FUNCTION_BLOCK FB_CIP EXTENDS FB_SFC_Cycle IMPLEMENTS ITF_FB_SFC_Cycle
VAR_INPUT
	valFillWater_T91	: E_Pis_Name;
	valFillWater_T92	: E_Pis_Name;
	valFillWater_T93	: E_Pis_Name;
	valFillWater_T94	: E_Pis_Name;
	
	lvlTank_T91			: ST_Tank_Level	;
	lvlTank_T92			: ST_Tank_Level	;
	lvlTank_T93			: ST_Tank_Level	;
	lvlTank_T94			: ST_Tank_Level	;

END_VAR
VAR_OUTPUT
END_VAR
VAR
	//bRun: BOOL;
	eRun: E_CIP_Source;

	eMode			: E_CIP_Mode;
	eCIP_Return		: E_CIP_Return;
	eCIP_Source		: E_CIP_Source;
	eCIP_Usage		: E_CIP_Usage;
	eReq			: ST_CIP_Request;
	eReqBlank		: ST_CIP_Request;
	eReqLocal		: ST_CIP_Request;
	
	ref_lvlTank_Client		: REFERENCE TO ST_Tank_Level	;

	//bStepDone: BOOL;
	
	iPosSelect_HMI: INT;

	rtPosMoveHMI_Up		: R_TRIG;
	rtPosMoveHMI_Down	: R_TRIG;
	rtPosDeleteHMI		: R_TRIG;
	rtPosDeleteAllHMI	: R_TRIG;
	
	eRefClient_fbElement		: REFERENCE TO FB_Element; // FB_Element // E_Element_State_Long
	bClientRef_done				: BOOL;
	fbElement_Blank				: FB_Element;
	eState_Long_Blank			: E_Element_State_Long;
	
	fbPis						: FB_Piston;
	stPis_FillWater_T91			: REFERENCE TO ST_Piston;
	stPis_FillWater_T92			: REFERENCE TO ST_Piston;
	stPis_FillWater_T93			: REFERENCE TO ST_Piston;
	stPis_FillWater_T94			: REFERENCE TO ST_Piston;
	
	rtReqLocalCIP_Full_HMI: R_TRIG;
	rtReqLocalCIP_Detergent_HMI: R_TRIG;
	rtReqCleanEmpty_HMI: R_TRIG;
	rtModeOff: R_TRIG;
	rtModeManual: R_TRIG;
	rtModeAuto: R_TRIG;
	bTemp: BOOL;
		
	//Process Control
	//concentration
	stDetergent					:	REFERENCE TO ST_ProcessControl	;
	pcDetergent					: 	REFERENCE TO FB_ProcessControl	;	//detergent local
	stDisInfectant				:	REFERENCE TO ST_ProcessControl	;
	pcDisInfectant				: 	REFERENCE TO FB_ProcessControl	;	//detergent local
    //temperature
	stHeatExchanger					:	REFERENCE TO ST_ProcessControl	;
	pcHeatExchanger					: 	REFERENCE TO FB_ProcessControl	;	//	
	stTemperature_Deterg			:	REFERENCE TO ST_ProcessControl	;
	pcTemperature_Deterg			: 	REFERENCE TO FB_ProcessControl	;	//detergent Client	
	stTemperature_Dis				:	REFERENCE TO ST_ProcessControl	;
	pcTemperature_Dis				: 	REFERENCE TO FB_ProcessControl	;//disinfectant local/client
	//temperature client return
	stTemp_ClntReturn				:	REFERENCE TO ST_ProcessControl	;//Client return temperature
	pcTemp_ClntReturn				: 	REFERENCE TO FB_ProcessControl	;//Client return temperature
	
	//flow rate
	stFlow1_Rate					:	REFERENCE TO ST_ProcessControl	;//CIP
	pcFlow1_Rate					: 	REFERENCE TO FB_ProcessControl	;//disinfectant local/client
	stFlow2_Rate					:	REFERENCE TO ST_ProcessControl	;//CIP send
	pcFlow2_Rate					: 	REFERENCE TO FB_ProcessControl	;//disinfectant local/client	return 
	stFlow3_Rate					:	REFERENCE TO ST_ProcessControl	;//CIP send
	pcFlow3_Rate					: 	REFERENCE TO FB_ProcessControl	;//disinfectant local/client	return 
	
	stColor_Level					:	REFERENCE TO ST_ProcessControl	;//CLient CIP //level control 
	pcColor_Level					: 	REFERENCE TO FB_ProcessControl	;//disinfectant local/client //level control 
	stMarinada_Level				:	REFERENCE TO ST_ProcessControl	;//CLient CIP //level control 
	pcMarinada_Level				: 	REFERENCE TO FB_ProcessControl	;//disinfectant local/client //level control 
	
	
	//colar marinade 
	//pressure
	stP1001_Pressure				:	REFERENCE TO ST_ProcessControl	;
	pcP1001_Pressure				: 	REFERENCE TO FB_ProcessControl	;//CIP //Client
(*
	stP3001_Pressure				:	REFERENCE TO ST_ProcessControl	;
	pcP3001_Pressure				: 	REFERENCE TO FB_ProcessControl	;
	
	stP3002_Pressure				:	REFERENCE TO ST_ProcessControl	;
	pcP3002_Pressure				: 	REFERENCE TO FB_ProcessControl	;	
	
	stP4001_Pressure				:	REFERENCE TO ST_ProcessControl	;
	pcP4001_Pressure				: 	REFERENCE TO FB_ProcessControl	;
	
	stP4002_Pressure				:	REFERENCE TO ST_ProcessControl	;
	pcP4002_Pressure				: 	REFERENCE TO FB_ProcessControl	;	
	
	stTriBlender_Flow				:	REFERENCE TO ST_ProcessControl	;
	pcTriBlender_Flow				: 	REFERENCE TO FB_ProcessControl	;	
	
	stColor_TriB_Conc				:	REFERENCE TO ST_ProcessControl	;
	pcColor_TriB_Conc				: 	REFERENCE TO FB_ProcessControl	;	
	
	stColor_Line_Conc				:	REFERENCE TO ST_ProcessControl	;
	pcColor_Line_Conc				: 	REFERENCE TO FB_ProcessControl	;	
*)	
	
		//OldOne to be deleted
		iStepDone: INT;
		fDetergTarget: REAL:=0.7;
		fDetergDeviation: REAL;
		fDetergLowTolerance: LREAL;
		fDetergHighTolerance: LREAL;
	

	
	bCIP_Condition_Failed: BOOL;
	testTemperature: REAL := 26.0;
	tonr_CIP_Condition: TONR;
	bCIP_Condition_Done: BOOL;
	fReqVolumeT93: REAL := 250;
	delta_T91_Volume: REAL;	// DisInfection
	delta_T92_Volume: REAL;	// Detergent
	delta_T93_Volume: REAL;	// Recycle Water
	delta_T94_Volume: REAL;	// Water
	memo_T91_Level_start: REAL;
	memo_T92_Level_start: REAL;
	memo_T93_Level_start: REAL;
	memo_T94_Level_start: REAL;	
	
	nStepHeat	:	INT		;
	
	bTestPID: BOOL;
	st_CIP_Param		:	ST_CIP_Param	;
	hystCIP_SetPoint: FB_Hysteresis_REAL;
	a: REAL := 0.8;
	b: REAL := 1.2;
	i: E_CIP_Usage;
	tMeasureDelayTime: TIME;
	bLoadDefSetPoints: BOOL;


	
	//Additional water valume if the solution concentration is too high
	rDeltaWater_DeterLocal		:	REAL	;
	rDeltaWater_DeterClient		:	REAL	;
	rDeltaWater_DisInfLocal		:	REAL	;
	rDeltaWater_DisInfClient	:	REAL	;

	rDeluteVolume				: REAL;
	rDeluteVolume_max			: REAL:=900;

	//accumulative actual time for desinfection and detergent condition
	nDeter_CondActTime_Lcl		:	INT	;//Actual condition time in seconds, for local client, detergent
	nDeter_CondActTime_Clnt		:	INT	;//Actual condition time in seconds, for client, detergent
	nDisInf_CondActTime_Lcl		:	INT	;//Actual condition time in seconds, for local client, disinfection
	nDisInf_CondActTime_Clnt	:	INT	;//Actual condition time in seconds, for client, disinfection
	
	bDeter_CondActTime_Lcl_Done		:	BOOL	;
	bDeter_CondActTime_Clnt_Done	:	BOOL	;
	bDisInf_CondActTime_Lcl_Done	:	BOOL	;
	bDisInf_CondActTime_Clnt_Done	:	BOOL	;

	fbHysteresisFillT94: FB_Hysteresis_REAL;
	
	//Choose pipe or sprinkler
	bSprinkler			:	BOOL:=FALSE	;
	tConditionTime		:	INT		;
	//tConditionTemper:	REAL	;
	fFlowRate			:	REAL	;
	//rVolume_Collect	:	REAL	;
	//rVolume_Drain		:	REAL	;
	//rVolume_Recycle	:	REAL	;
	
	_temp: REAL;
	_cond: ARRAY[0..9] OF BOOL;
	tonStepConditionTime: TON;
	bClientTypeIs_Tank: BOOL;
	t_ActMeasureTime: TIME;
	
	volume_Requered	: INT;
	volume_Actual	: INT;

	ton_Concentration_Filter: TON;
	bConcentration_correct: BOOL;
	tonTankLowLevel: TON;
	iCheck: INT;
	bMixProof_Release_All: BOOL;
	iConcentrationDeluteCounter: INT;
END_VAR
//upper lower control
VAR
	nClient			:	INT:=1		;
	bClean_MixProof	:	BOOL:=FALSE	;
	nNumOfRetries	:	INT:=5		;
	nNumOfPulses	:	INT:=5		;//Number of pulses per valve seat clean
	nStep_Vlv		:	INT:=0		;
	bValveCleanDone	:	BOOL:=FALSE	;
	nI_1_act_valve			:	INT:=1		;
	nI_2_act_pulses			:	INT:=0		;
	nI_3_act_repeats		:	INT:=1		;//number of repeats
	ActvValve		:	E_Pis_Name	;
	bSeatStatus		:	BOOL:=FALSE	;
	sState			:	STRING		;
	tOn				:	TON			;
	tOff			:	TON			;
	
	nMaxValves		:	INT:=6		;
	
	arTestOverflow: ARRAY[0..5] OF REAL;

END_VAR

VAR_IN_OUT
	fbCIP_Source	: FB_CIP_Source	;
	fbCIP_Return	: FB_CIP_Return	;
	fbCIP_Usage		: FB_CIP_Client	;
	
	//fbTarget					: FB_Tank_Target	;
	//fbLineSource				: FB_Line_Source	;
	//fbLineTarget				: FB_Line_Target	;
	//fbTriBlenderSource		: FB_Line_Source	;
	//fbTriBlenderTarget		: FB_Line_Target	;

	//fb_PumpLine				: FB_Pump	;
	//fb_PumpTriBlender			: FB_Pump	;
	fbTank1	:	FB_ProductionTank	;
	fbTank2	:	FB_ProductionTank	;
	fbTank3	:	FB_ProductionTank	;
	fbTank4	:	FB_ProductionTank	;
	
	//Pumps
	fb_PumpCIP				: FB_Pump;
	fb_PumpClient			: FB_Pump;
	fb_Stirrer				: FB_Pump;
	fb_PumpDetergent		: FB_DosingPump;
	fb_PumpDisinfection		: FB_DosingPump;
	
	//Heat Exchenger	
	fb_HeatExchenger	:	FB_HeatExchanger	;
	

END_VAR

m_Set_SFCFlags_Reference();
act_GetReference();
act_CallProcessControl();
//act_HeatExchng();
act_SprinklerCondition();
//SUPER^();

//Selecting client for CIP parameters
st_CIP_Param:=g_Data.arr_CIP_Param[eReq.eClient];
FOR i:=1 TO E_CIP_Usage.eLocal DO
	g_Data.arr_CIP_Param[i].sName:=TO_STRING(i);
END_FOR

act_Oper();
act_ReqBuffer();
mVolumeMeter();
act_ValveUpLow_Cntrl();

rtModeOff(CLK:=eMode=E_CIP_Mode.eOff);
IF rtModeOff.Q THEN;
	SFCReset:=TRUE;
END_IF

rtModeManual(CLK:=eMode=E_CIP_Mode.eManual);
IF rtModeManual.Q THEN;
	bTemp:=TRUE;
END_IF

rtModeAuto(CLK:=eMode=E_CIP_Mode.eAuto);
IF rtModeAuto.Q THEN;
	//SFCReset:=TRUE;
END_IF

IF bRun AND bClientRef_done THEN;
	act_Run();
END_IF


t_ActMeasureTime:=m_MeasureTimeToHMI();
mFillWater();
//IF bMoveStep THEN bMoveStep:=FALSE; END_IF
IF bMixProof_Release_All THEN;
	IF m_MixProof_Release_All() THEN;
		bMixProof_Release_All:=FALSE;
	END_IF
END_IF
m_DashState_MixProof_set();
(*
arTestOverflow[0]:=m_OverFlowCorrect(
rTc:=arTestOverflow[1], 
rAv:=arTestOverflow[2], 
rAc:=arTestOverflow[3]);
*)

ACTION _aCIP1_Conn_Sprinkler_active:
//Connect client tank to sprinkler
CASE eReq.eClient OF
	
	E_CIP_Usage.eTank_1:;
				bStepDone:=fbCIP_ClientTank_Marinade.m_CheckStatus(eReqStatus:=E_CIP_ClientTank.eTank_A_Sprinkler);
	E_CIP_Usage.eTank_2:;
				bStepDone:=fbCIP_ClientTank_Marinade.m_CheckStatus(eReqStatus:=E_CIP_ClientTank.eTank_B_Sprinkler);	
	E_CIP_Usage.eTank_3:;
				bStepDone:=fbCIP_ClientTank_Color.m_CheckStatus(eReqStatus:=E_CIP_ClientTank.eTank_A_Sprinkler);
	E_CIP_Usage.eTank_4:;
				bStepDone:=fbCIP_ClientTank_Color.m_CheckStatus(eReqStatus:=E_CIP_ClientTank.eTank_B_Sprinkler);	

ELSE;				
	bStepDone:=FALSE;
END_CASE
END_ACTION

ACTION _aCIP1_Conn_Sprinkler_entry:
bSprinkler:=TRUE;
CASE eReq.eClient OF

	E_CIP_Usage.eTank_1:;
				fbCIP_ClientTank_Marinade.m_Run(eReqProc:=E_CIP_ClientTank.eTank_A_Sprinkler);
	E_CIP_Usage.eTank_2:;
				fbCIP_ClientTank_Marinade.m_Run(eReqProc:=E_CIP_ClientTank.eTank_B_Sprinkler);	
	E_CIP_Usage.eTank_3:;
				fbCIP_ClientTank_Color.m_Run(eReqProc:=E_CIP_ClientTank.eTank_A_Sprinkler);
	E_CIP_Usage.eTank_4:;
				fbCIP_ClientTank_Color.m_Run(eReqProc:=E_CIP_ClientTank.eTank_B_Sprinkler);	

END_CASE
tonr_CIP_Condition(ResetTime:=TRUE);
END_ACTION

ACTION _aCIP1_Done_entry:
eRefClient_fbElement.m_InterConnected_State(eState_Long_Set:=E_Element_State_Long.eCIP_1_Rinzed);
END_ACTION

ACTION _aCIP2_Conn_Sprinkler_active:
//Connect client tank to sprinkler
CASE eReq.eClient OF
	
	E_CIP_Usage.eTank_1:;
				bStepDone:=fbCIP_ClientTank_Marinade.m_CheckStatus(eReqStatus:=E_CIP_ClientTank.eTank_A_Sprinkler);
	E_CIP_Usage.eTank_2:;
				bStepDone:=fbCIP_ClientTank_Marinade.m_CheckStatus(eReqStatus:=E_CIP_ClientTank.eTank_B_Sprinkler);	
	E_CIP_Usage.eTank_3:;
				bStepDone:=fbCIP_ClientTank_Color.m_CheckStatus(eReqStatus:=E_CIP_ClientTank.eTank_A_Sprinkler);
	E_CIP_Usage.eTank_4:;
				bStepDone:=fbCIP_ClientTank_Color.m_CheckStatus(eReqStatus:=E_CIP_ClientTank.eTank_B_Sprinkler);	

ELSE;				
	bStepDone:=FALSE;
END_CASE
END_ACTION

ACTION _aCIP2_Conn_Sprinkler_entry:
//bSprinkler:=TRUE;
CASE eReq.eClient OF

	E_CIP_Usage.eTank_1:;
				fbCIP_ClientTank_Marinade.m_Run(eReqProc:=E_CIP_ClientTank.eTank_A_Sprinkler);
	E_CIP_Usage.eTank_2:;
				fbCIP_ClientTank_Marinade.m_Run(eReqProc:=E_CIP_ClientTank.eTank_B_Sprinkler);	
	E_CIP_Usage.eTank_3:;
				fbCIP_ClientTank_Color.m_Run(eReqProc:=E_CIP_ClientTank.eTank_A_Sprinkler);
	E_CIP_Usage.eTank_4:;
				fbCIP_ClientTank_Color.m_Run(eReqProc:=E_CIP_ClientTank.eTank_B_Sprinkler);	

END_CASE
tonr_CIP_Condition(ResetTime:=TRUE);
END_ACTION

ACTION _aCIP2_Done_entry:
IF eReq.eClient=E_CIP_Usage.eLocal THEN;
	eRefClient_fbElement.m_InterConnected_State(eState_Long_Set:=E_Element_State_Long.eCIP_2_Deterged);
ELSE;
	eRefClient_fbElement.m_InterConnected_State(eState_Long_Set:=E_Element_State_Long.eCIP_2_Deterged);
END_IF
END_ACTION

ACTION _aCIP2_Flow_Sprincler_active:
fb_PumpCIP.m_Run(RPM:=pcFlow1_Rate.mRun_PID(Set_Point:=fFlowRate, controlManual:=NOT(fb_PumpCIP.modeAuto)));
fb_PumpClient.m_Run(RPM:=st_CIP_Param.r_CIP_Client_Pump);

IF TRUE 
AND pcFlow1_Rate.mRun()
AND pcFlow2_Rate.mRun()
//AND pcPressure.mRun()
THEN;
	tonStepConditionTime.IN:=TRUE;
ELSE;
	tonStepConditionTime.IN:=FALSE;
END_IF

tonStepConditionTime(PT:=T#10S);
IF tonStepConditionTime.Q THEN;
	bStepDone:=TRUE;
ELSE;
	bStepDone:=FALSE;
END_IF
END_ACTION

ACTION _aCIP2_Flow_Sprincler_entry:
tonStepConditionTime(IN:=FALSE);

m_DashState_done(stage:=E_CIP_DashStage_List.e06_CIP2_Client_Detergent_Condition_Pipe);
m_DashState_activate(stage:=E_CIP_DashStage_List.e07_CIP2_Client_Detergent_Condition_Sprinkler);
END_ACTION

ACTION _aCIP2_If_ClientIsTank_active:
CASE eReq.eClient OF
	E_CIP_Usage.eTank_1,
	E_CIP_Usage.eTank_2,
	E_CIP_Usage.eTank_3,
	E_CIP_Usage.eTank_4:;
			bStepDone:=TRUE;
			m_DashState_done(stage:=E_CIP_DashStage_List.e07_CIP2_Client_Detergent_Condition_Sprinkler);
			
ELSE;
			bStepDone:=FALSE;
			m_DashState_done(stage:=E_CIP_DashStage_List.e06_CIP2_Client_Detergent_Condition_Pipe);
END_CASE
END_ACTION

ACTION _aCIP3_Conn_Sprinkler_active:
//Connect client tank to sprinkler
CASE eReq.eClient OF
	
	E_CIP_Usage.eTank_1:;
				bStepDone:=fbCIP_ClientTank_Marinade.m_CheckStatus(eReqStatus:=E_CIP_ClientTank.eTank_A_Sprinkler);
	E_CIP_Usage.eTank_2:;
				bStepDone:=fbCIP_ClientTank_Marinade.m_CheckStatus(eReqStatus:=E_CIP_ClientTank.eTank_B_Sprinkler);	
	E_CIP_Usage.eTank_3:;
				bStepDone:=fbCIP_ClientTank_Color.m_CheckStatus(eReqStatus:=E_CIP_ClientTank.eTank_A_Sprinkler);
	E_CIP_Usage.eTank_4:;
				bStepDone:=fbCIP_ClientTank_Color.m_CheckStatus(eReqStatus:=E_CIP_ClientTank.eTank_B_Sprinkler);	
ELSE;				
	bStepDone:=FALSE;
END_CASE
END_ACTION

ACTION _aCIP3_Conn_Sprinkler_entry:
//bSprinkler:=TRUE;
CASE eReq.eClient OF

	E_CIP_Usage.eTank_1:;
				fbCIP_ClientTank_Marinade.m_Run(eReqProc:=E_CIP_ClientTank.eTank_A_Sprinkler);
	E_CIP_Usage.eTank_2:;
				fbCIP_ClientTank_Marinade.m_Run(eReqProc:=E_CIP_ClientTank.eTank_B_Sprinkler);	
	E_CIP_Usage.eTank_3:;
				fbCIP_ClientTank_Color.m_Run(eReqProc:=E_CIP_ClientTank.eTank_A_Sprinkler);
	E_CIP_Usage.eTank_4:;
				fbCIP_ClientTank_Color.m_Run(eReqProc:=E_CIP_ClientTank.eTank_B_Sprinkler);	

END_CASE
tonr_CIP_Condition(ResetTime:=TRUE);
END_ACTION

ACTION _aCIP3_Done_entry:
eRefClient_fbElement.m_InterConnected_State(eState_Long_Set:=E_Element_State_Long.eCIP_4_Sanitized);
END_ACTION

ACTION _aCIP3_Flow_Sprincler_active:
fb_PumpCIP.m_Run(RPM:=pcFlow1_Rate.mRun_PID(Set_Point:=fFlowRate, controlManual:=NOT(fb_PumpCIP.modeAuto)));
fb_PumpClient.m_Run(RPM:=st_CIP_Param.r_CIP_Client_Pump);

IF TRUE 
AND pcFlow1_Rate.mRun()
AND pcFlow2_Rate.mRun()
//AND pcPressure.mRun()
THEN;
	tonStepConditionTime.IN:=TRUE;
ELSE;
	tonStepConditionTime.IN:=FALSE;
END_IF

tonStepConditionTime(PT:=T#10S);
IF tonStepConditionTime.Q THEN;
	bStepDone:=TRUE;
ELSE;
	bStepDone:=FALSE;
END_IF
END_ACTION

ACTION _aCIP3_Flow_Sprincler_entry:
tonStepConditionTime(IN:=FALSE);
m_DashState_done(stage:=E_CIP_DashStage_List.e15_CIP4_Client_DisInfection_Condition_Pipe);
m_DashState_activate(stage:=E_CIP_DashStage_List.e16_CIP4_Client_DisInfection_Condition_Sprinkler);
END_ACTION

ACTION _aCIP3_If_ClientIsTank_active:
CASE eReq.eClient OF
	E_CIP_Usage.eTank_1,
	E_CIP_Usage.eTank_2,
	E_CIP_Usage.eTank_3,
	E_CIP_Usage.eTank_4:;
		bStepDone:=TRUE;
		m_DashState_done(stage:=E_CIP_DashStage_List.e16_CIP4_Client_DisInfection_Condition_Sprinkler);
ELSE;
		bStepDone:=FALSE;
		m_DashState_done(stage:=E_CIP_DashStage_List.e15_CIP4_Client_DisInfection_Condition_Pipe);
END_CASE
END_ACTION

ACTION _aCIP4_Collect_active:
bStepDone:=FALSE;
IF eRefClient_fbElement.eState_Long=E_Element_State_Long.eCIP_2_Deterged THEN;
	volume_Requered:= REAL_TO_INT(st_CIP_Param.r_Volume_Collect_Detergent);
	volume_Actual:= REAL_TO_INT(delta_T92_Volume);
ELSIF eRefClient_fbElement.eState_Long=E_Element_State_Long.eCIP_4_Sanitized THEN;
	volume_Requered:= REAL_TO_INT(st_CIP_Param.r_Volume_Collect_DisInfection);
	volume_Actual:= REAL_TO_INT(delta_T91_Volume);
END_IF

IF volume_Actual >= volume_Requered THEN;
	bStepDone:=TRUE;
END_IF

(*
IF TRUE 
OR (delta_T94_Volume < -st_CIP_Param.r_Volume_Collect_Detergent AND eRefClient_fbElement.eState_Long=E_Element_State_Long.eCIP_2_Deterged)
OR (delta_T94_Volume < -st_CIP_Param.r_Volume_Collect_DisInfection AND eRefClient_fbElement.eState_Long=E_Element_State_Long.eCIP_4_Sanitized)

OR (delta_T92_Volume > st_CIP_Param.r_Volume_Collect_Detergent AND eRefClient_fbElement.eState_Long=E_Element_State_Long.eCIP_2_Deterged)
OR (delta_T91_Volume > st_CIP_Param.r_Volume_Collect_DisInfection AND eRefClient_fbElement.eState_Long=E_Element_State_Long.eCIP_4_Sanitized)
THEN
	bStepDone:=TRUE;
END_IF
*)
END_ACTION

ACTION _aCIP4_Collect_entry:
mVolumeReset_All();
END_ACTION

ACTION _aCIP4_Conn_Sprinkler_active:
//Connect client tank to sprinkler
CASE eReq.eClient OF
	
	E_CIP_Usage.eTank_1:;
				bStepDone:=fbCIP_ClientTank_Marinade.m_CheckStatus(eReqStatus:=E_CIP_ClientTank.eTank_A_Sprinkler);
	E_CIP_Usage.eTank_2:;
				bStepDone:=fbCIP_ClientTank_Marinade.m_CheckStatus(eReqStatus:=E_CIP_ClientTank.eTank_B_Sprinkler);	
	E_CIP_Usage.eTank_3:;
				bStepDone:=fbCIP_ClientTank_Color.m_CheckStatus(eReqStatus:=E_CIP_ClientTank.eTank_A_Sprinkler);
	E_CIP_Usage.eTank_4:;
				bStepDone:=fbCIP_ClientTank_Color.m_CheckStatus(eReqStatus:=E_CIP_ClientTank.eTank_B_Sprinkler);	

ELSE;				
	bStepDone:=FALSE;
END_CASE
END_ACTION

ACTION _aCIP4_Conn_Sprinkler_entry:
bSprinkler:=TRUE;
CASE eReq.eClient OF

	E_CIP_Usage.eTank_1:;
				fbCIP_ClientTank_Marinade.m_Run(eReqProc:=E_CIP_ClientTank.eTank_A_Sprinkler);
	E_CIP_Usage.eTank_2:;
				fbCIP_ClientTank_Marinade.m_Run(eReqProc:=E_CIP_ClientTank.eTank_B_Sprinkler);	
	E_CIP_Usage.eTank_3:;
				fbCIP_ClientTank_Color.m_Run(eReqProc:=E_CIP_ClientTank.eTank_A_Sprinkler);
	E_CIP_Usage.eTank_4:;
				fbCIP_ClientTank_Color.m_Run(eReqProc:=E_CIP_ClientTank.eTank_B_Sprinkler);	

END_CASE
tonr_CIP_Condition(ResetTime:=TRUE);
END_ACTION

ACTION _aCIP4_Done_entry:


CASE eRefClient_fbElement.eState_Long OF
	E_Element_State_Long.eNotClean:;
			//
	E_Element_State_Long.eCIP_1_Rinzed:;
			//
	E_Element_State_Long.eCIP_2_Deterged:;
			eRefClient_fbElement.m_InterConnected_State(eState_Long_Set:=E_Element_State_Long.eCIP_3_Deterged_Clean);	
		
	E_Element_State_Long.eCIP_3_Deterged_Clean:;
			//
	E_Element_State_Long.eCIP_4_Sanitized:;
			eRefClient_fbElement.m_InterConnected_State(eState_Long_Set:=E_Element_State_Long.eCIP_5_Done);			
	
END_CASE
END_ACTION

ACTION _aCIP4_Drain_active:
bStepDone:=FALSE;

IF eRefClient_fbElement.eState_Long=E_Element_State_Long.eCIP_2_Deterged THEN;
	volume_Requered:= REAL_TO_INT(st_CIP_Param.r_Volume_Drain_Detergent);
	volume_Actual:= REAL_TO_INT(-delta_T94_Volume);
ELSIF eRefClient_fbElement.eState_Long=E_Element_State_Long.eCIP_4_Sanitized THEN;
	volume_Requered:= REAL_TO_INT(st_CIP_Param.r_Volume_Drain_DisInfection);
	volume_Actual:= REAL_TO_INT(-delta_T94_Volume);
END_IF

IF volume_Actual >= volume_Requered THEN;
	bStepDone:=TRUE;
END_IF


(*
IF fbCIP_Return.m_CheckStatus(eReqStatus:=E_CIP_Return.eDrain)  
AND ((delta_T94_Volume < -st_CIP_Param.r_Volume_Drain_Detergent AND eRefClient_fbElement.eState_Long=E_Element_State_Long.eCIP_2_Deterged)
OR (delta_T94_Volume < -st_CIP_Param.r_Volume_Drain_DisInfection AND eRefClient_fbElement.eState_Long=E_Element_State_Long.eCIP_4_Sanitized))
//TEMP T93
//OR (delta_T93_Volume < -st_CIP_Param.r_Volume_Drain_Detergent AND eRefClient_fbElement.eState_Long=E_Element_State_Long.eCIP_2_Deterged)
//OR (delta_T93_Volume < -st_CIP_Param.r_Volume_Drain_DisInfection AND eRefClient_fbElement.eState_Long=E_Element_State_Long.eCIP_4_Sanitized))
THEN;
	bStepDone:=TRUE;
END_IF
*)
END_ACTION

ACTION _aCIP4_Drain_entry:
fbCIP_Return.m_Run(eReqProc:=E_CIP_Return.eDrain);
mVolumeReset_All();

CASE eRefClient_fbElement.eState_Long OF

	E_Element_State_Long.eCIP_2_Deterged:;
			m_DashState_done(stage:=E_CIP_DashStage_List.e08_CIP3_Detergent_Collect);
			m_DashState_activate(stage:=E_CIP_DashStage_List.e09_CIP3_Detergent_Drain);

	E_Element_State_Long.eCIP_4_Sanitized:;
			m_DashState_done(stage:=E_CIP_DashStage_List.e17_CIP5_DisInfection_Collect);
			m_DashState_activate(stage:=E_CIP_DashStage_List.e18_CIP5_DisInfection_Drain);
			
END_CASE
END_ACTION

ACTION _aClient_tank_IsEmpty_active:
bStepDone:=m_ClientTank_IsEmpty();

(*
IF bClientTypeIs_Tank THEN;
	//
END_IF
CASE eCIP_Usage OF
	E_CIP_Usage.eTank_1:;
			IF stTanksSens[E_Tank_Name.T1].e_state=E_Tank_Level.eEmpty THEN;
				bStepDone:=TRUE;	
			END_IF	
	E_CIP_Usage.eTank_2:;
			IF stTanksSens[E_Tank_Name.T2].e_state=E_Tank_Level.eEmpty THEN;
				bStepDone:=TRUE;	
			END_IF	
	E_CIP_Usage.eTank_3:;
			IF stTanksSens[E_Tank_Name.T3].e_state=E_Tank_Level.eEmpty THEN;
				bStepDone:=TRUE;	
			END_IF	
	E_CIP_Usage.eTank_4:;
			IF stTanksSens[E_Tank_Name.T4].e_state=E_Tank_Level.eEmpty THEN;
				bStepDone:=TRUE;	
			END_IF
ELSE;
	bStepDone:=TRUE;	
END_CASE
*)
END_ACTION

ACTION _aClient_Validation_check_active:
bStepDone:=FALSE;
	
IF eRefClient_fbElement.m_Get_Type()=E_Element_Type.eTriBlender THEN;
	IF TRUE 
	AND fbElement[E_Element_List.eTriBlender_Color].m_Get_CIP_Avilable()
	AND fbElement[E_Element_List.eTriBlender_Marinada].m_Get_CIP_Avilable()
	AND eRun<>E_CIP_Source.eNone
	AND TRUE
	THEN;
		bStepDone:=eRefClient_fbElement.m_InterConnect(value:=E_InterConnection.ConnToCIP);		
	END_IF		
ELSE;
	IF TRUE 
	AND eRefClient_fbElement.m_Get_CIP_Avilable()
	AND eRun<>E_CIP_Source.eNone
	AND TRUE
	THEN;
		bStepDone:=eRefClient_fbElement.m_InterConnect(value:=E_InterConnection.ConnToCIP);
	END_IF
END_IF
END_ACTION

ACTION _aClientReference_IsValid_entry:
IF bClientTypeIs_Tank THEN;
	fb_Stirrer.m_Run(RPM:=1200);
END_IF
END_ACTION

ACTION _aCondition_CIP1_Client_active:
IF NOT bSprinkler THEN
	//pipe
	tConditionTime	:=st_CIP_Param.t_ConditionR_Water;
	fFlowRate		:=st_CIP_Param.r_Flow_Pipe;
	
ELSE
	//sprinkler
	tConditionTime	:=st_CIP_Param.t_ConditionR_Water_Sprinkler;
	fFlowRate		:=st_CIP_Param.r_Flow_Sprinkler;
END_IF

IF Condition_CIP1_Client.t > SECOND_TO_TIME(st_CIP_Param.t_PumpInitRun) THEN;
	fb_PumpCIP.m_Run(RPM:=pcFlow1_Rate.mRun_PID(Set_Point:=fFlowRate,controlManual:=NOT(fb_PumpCIP.modeAuto)));
END_IF


tonr_CIP_Condition(PT:=SECOND_TO_TIME(tConditionTime));
//
IF bSprinkler THEN;
	IF TRUE 
	AND pcFlow1_Rate.mRun(mRun=>_cond[1])
	//AND pcFlow3_Rate.mRun(mRun=>_cond[2])
	THEN;
		tonr_CIP_Condition.IN:=TRUE;
	ELSE;
		tonr_CIP_Condition.IN:=FALSE;
	END_IF
ELSE;
	IF TRUE 
	AND pcFlow1_Rate.mRun(mRun=>_cond[1])
	//AND pcFlow2_Rate.mRun(mRun=>_cond[2])
	THEN;
		tonr_CIP_Condition.IN:=TRUE;
	ELSE;
		tonr_CIP_Condition.IN:=FALSE;
	END_IF	
	
END_IF
//

IF tonr_CIP_Condition.Q THEN
	bCIP_Condition_Done:=TRUE;
ELSE;
	bCIP_Condition_Done:=FALSE;	
END_IF

IF FALSE  
//AND delta_T93_Volume < -st_CIP_Param.r_Volume_Drain_R_Water 
OR lvlTank_T93.rTankLevel < 250
THEN;
	bCIP_Condition_Failed:=TRUE;
END_IF



(*
// Connect return to R_Water
IF TRUE 
AND lvlTank_T93.rTankLevel<450 
AND fbCIP_Return.m_CheckStatus(eReqStatus:=E_CIP_Return.eDrain)
THEN;
	fbCIP_Return.m_Run(eReqProc:=E_CIP_Return.eT93_R_Water);
ELSE;
	
END_IF



// Connect return to Drain

IF TRUE 
AND lvlTank_T93.rTankLevel>500 // The tank is full
AND fbCIP_Return.m_CheckStatus(eReqStatus:=E_CIP_Return.eT93_R_Water)
THEN;
	fbCIP_Return.m_Run(eReqProc:=E_CIP_Return.eDrain);
ELSE;
	
END_IF
*)


(*
IF TRUE 
AND bCIP_Condition_Done
OR bCIP_Condition_Failed
THEN;

ELSE;
	
END_IF

IF TRUE 
AND pcFlow1_Rate.mRun(mRun=>_cond[1])
AND pcFlow2_Rate.mRun(mRun=>_cond[2])
//AND pcPressure.mRun()
THEN;
	//
ELSE;
	bCIP_Condition_Failed:=TRUE;
END_IF
*)
END_ACTION

ACTION _aCondition_CIP1_Client_entry:
//fbCIP_Return.m_Run(eReqProc:=E_CIP_Return.eT93_R_Water);

fb_PumpCIP.m_Run(RPM:=st_CIP_Param.r_CIP_Pump);
fb_PumpClient.m_Run(RPM:=st_CIP_Param.r_CIP_Client_Pump);

bCIP_Condition_Failed:=FALSE;
bCIP_Condition_Done:=FALSE;
mVolumeReset_All();
END_ACTION

ACTION _aCondition_CIP1_Client_exit:
tonr_CIP_Condition(IN:=FALSE);
END_ACTION

ACTION _aCondition_CIP2_Client_active:
fb_PumpCIP.m_Run(RPM:=pcFlow1_Rate.mRun_PID(Set_Point:=fFlowRate, controlManual:=NOT(fb_PumpCIP.modeAuto)));
fb_PumpClient.m_Run(RPM:=st_CIP_Param.r_CIP_Client_Pump);

IF bSprinkler THEN;
	IF TRUE 
	AND pcFlow1_Rate.mRun(mRun=>_cond[1])
	AND pcFlow3_Rate.mRun(mRun=>_cond[2])
	THEN;
		//
	ELSE;
		bCIP_Condition_Failed:=TRUE;
	END_IF
ELSE;
	IF TRUE 
	AND pcFlow1_Rate.mRun(mRun=>_cond[1])
	AND pcFlow2_Rate.mRun(mRun=>_cond[2])
	THEN;
		//
	ELSE;
		bCIP_Condition_Failed:=TRUE;
	END_IF	
END_IF

pcHeatExchanger.mRun_PID(Set_Point:=st_CIP_Param.r_Temper_Detergent, controlManual:=g_Data.stHeatExchanger.bManual ,mRun_PID=>_temp);
tonr_CIP_Condition(PT:=SECOND_TO_TIME(tConditionTime));
IF TRUE 
AND pcHeatExchanger.mRun_With_SP(Set_Point:=st_CIP_Param.r_Temper_Detergent, mRun_With_SP=>_cond[3])
//AND pcTemperature_Deterg.mRun_With_SP(Set_Point:=g_Data.arr_CIP_Param[E_CIP_Usage.eLocal].r_Temper_Detergent, mRun_With_SP=>_cond[4])
AND pcTemp_ClntReturn.mRun_With_SP(Set_Point:=st_CIP_Param.r_Temper_Detergent, mRun_With_SP=>_cond[5])
AND pcDetergent.mRun_With_SP(Set_Point:=st_CIP_Param.r_DetergentConcentration, mRun_With_SP=>_cond[6])
AND measure_Deterg_2.x
AND TRUE
THEN;
	tonr_CIP_Condition.IN:=TRUE;
	m_MixProof_run();
ELSE;
	tonr_CIP_Condition.IN:=FALSE;
END_IF

IF tonr_CIP_Condition.Q 
AND bValveCleanDone
THEN;
	bCIP_Condition_Done:=TRUE;
ELSE;
	bCIP_Condition_Done:=FALSE;
END_IF



ton_Concentration_Filter(PT:=T#30S, IN:=stDetergent.Control_ON AND NOT stDetergent.OverFlow);
IF TRUE 
AND ton_Concentration_Filter.Q	
THEN;
	bConcentration_correct:=TRUE;
ELSE;
	bConcentration_correct:=FALSE;
END_IF

// Reverce function
(*
IF Deterg_Conc_Client_Done.x 
AND NOT pcDetergent.mRun() 
THEN;
	bCIP_Condition_Failed:=TRUE;
END_IF

IF Temperature_2_Done.x 
//AND NOT pcTemperature_Deterg.mRun()
AND NOT pcTemp_ClntReturn.mRun()
THEN;
	bCIP_Condition_Failed:=TRUE;
END_IF
*)
(*
//ton_CIP_Condition(PT:=T#30S);
IF tConditionTime-nDeter_CondActTime_Clnt>0 THEN
	tonr_CIP_Condition(PT:=SECOND_TO_TIME(tConditionTime-nDeter_CondActTime_Clnt));
	bDeter_CondActTime_Clnt_Done:=FALSE;
ELSE
	bDeter_CondActTime_Clnt_Done:=TRUE;
END_IF

IF TRUE 
AND Deterg_Conc_Client_Done.x
AND Temperature_2_Done.x
AND NOT bDeter_CondActTime_Clnt_Done
AND TRUE
THEN;
	tonr_CIP_Condition.IN:=TRUE;
ELSE;
	nDeter_CondActTime_Clnt:=TIME_TO_INT(tonr_CIP_Condition.ET)/1000;
	tonr_CIP_Condition.IN:=FALSE;
END_IF

IF tonr_CIP_Condition.Q
OR bDeter_CondActTime_Clnt_Done THEN;
	bCIP_Condition_Done:=TRUE;
ELSE;
	bCIP_Condition_Done:=FALSE;
END_IF
*)
END_ACTION

ACTION _aCondition_CIP2_Client_exit:
tonr_CIP_Condition(IN:=FALSE);
END_ACTION

ACTION _aCondition_CIP2_Local_active:
fb_PumpCIP.m_Run(RPM:=pcFlow1_Rate.mRun_PID(Set_Point:=g_Data.arr_CIP_Param[E_CIP_Usage.eLocal].r_Flow_Pipe,controlManual:=NOT(fb_PumpCIP.modeAuto)));

IF TRUE 
AND pcFlow1_Rate.mRun(mRun=>_cond[1])
AND pcFlow2_Rate.mRun(mRun=>_cond[2])
//AND pcPressure.mRun()
THEN;
	//
ELSE;
	bCIP_Condition_Failed:=TRUE;
END_IF

pcHeatExchanger.mRun_PID(Set_Point:=g_Data.arr_CIP_Param[E_CIP_Usage.eLocal].r_Temper_Detergent, controlManual:=g_Data.stHeatExchanger.bManual ,mRun_PID=>_temp);
tonr_CIP_Condition(PT:=SECOND_TO_TIME(g_Data.arr_CIP_Param[E_CIP_Usage.eLocal].t_ConditionDetergent), ResetTime:=FALSE);
IF TRUE 
AND pcHeatExchanger.mRun_With_SP(Set_Point:=g_Data.arr_CIP_Param[E_CIP_Usage.eLocal].r_Temper_Detergent, mRun_With_SP=>_cond[3])
AND pcTemperature_Deterg.mRun_With_SP(Set_Point:=g_Data.arr_CIP_Param[E_CIP_Usage.eLocal].r_Temper_Detergent, mRun_With_SP=>_cond[4])
AND pcTemp_ClntReturn.mRun_With_SP(Set_Point:=g_Data.arr_CIP_Param[E_CIP_Usage.eLocal].r_Temper_Detergent, mRun_With_SP=>_cond[5])
AND pcDetergent.mRun_With_SP(Set_Point:=g_Data.arr_CIP_Param[E_CIP_Usage.eLocal].r_DetergentConcentration, mRun_With_SP=>_cond[6])
AND measure_Deterg.x
AND TRUE
THEN;
	tonr_CIP_Condition.IN:=TRUE;
ELSE;
	tonr_CIP_Condition.IN:=FALSE;
END_IF
	
IF tonr_CIP_Condition.Q THEN;
	bCIP_Condition_Done:=TRUE;
ELSE;
	bCIP_Condition_Done:=FALSE;	
END_IF


ton_Concentration_Filter(PT:=T#30S, IN:=stDetergent.Control_ON AND NOT stDetergent.OverFlow);
IF TRUE 
AND ton_Concentration_Filter.Q	
THEN;
	bConcentration_correct:=TRUE;
ELSE;
	bConcentration_correct:=FALSE;
END_IF

// Reverce function

(*
IF Deterg_Conc_Local_Done.x 
AND NOT pcDetergent.mRun()
THEN;
	bCIP_Condition_Failed:=TRUE;
END_IF

IF Temperature_1_Done.x 
AND (NOT pcTemperature_Deterg.mRun()
	OR NOT pcTemp_ClntReturn.mRun())
THEN;
	bCIP_Condition_Failed:=TRUE;
END_IF
*)

(*
//ton_CIP_Condition(PT:=T#30S);
IF (g_Data.arr_CIP_Param[E_CIP_Usage.eLocal].t_ConditionDetergent-nDeter_CondActTime_Lcl)>0 THEN
	tonr_CIP_Condition(PT:=SECOND_TO_TIME(g_Data.arr_CIP_Param[E_CIP_Usage.eLocal].t_ConditionDetergent-nDeter_CondActTime_Lcl));
	bDeter_CondActTime_Lcl_Done:=FALSE;
ELSE
	bDeter_CondActTime_Lcl_Done:=TRUE;
END_IF

IF TRUE 
AND Deterg_Conc_Local_Done.x
AND Temperature_1_Done.x
AND NOT bDeter_CondActTime_Lcl_Done
AND TRUE
THEN;
	tonr_CIP_Condition.IN:=TRUE;
ELSE;
	nDeter_CondActTime_Lcl:=TIME_TO_INT(tonr_CIP_Condition.ET)/1000;
	tonr_CIP_Condition.IN:=FALSE;
END_IF
	
IF tonr_CIP_Condition.Q OR bDeter_CondActTime_Lcl_Done THEN;
	bCIP_Condition_Done:=TRUE;
ELSE;
	bCIP_Condition_Done:=FALSE;	
END_IF

*)
END_ACTION

ACTION _aCondition_CIP2_Local_exit:
tonr_CIP_Condition(IN:=FALSE);
END_ACTION

ACTION _aCondition_CIP3_Client_active:
fb_PumpCIP.m_Run(RPM:=pcFlow1_Rate.mRun_PID(Set_Point:=fFlowRate,controlManual:=NOT(fb_PumpCIP.modeAuto)));
fb_PumpClient.m_Run(RPM:=st_CIP_Param.r_CIP_Client_Pump);

IF bSprinkler THEN;
	IF TRUE 
	AND pcFlow1_Rate.mRun(mRun=>_cond[1])
	AND pcFlow3_Rate.mRun(mRun=>_cond[2])
	THEN;
		//
	ELSE;
		bCIP_Condition_Failed:=TRUE;
	END_IF
ELSE;
	IF TRUE 
	AND pcFlow1_Rate.mRun(mRun=>_cond[1])
	AND pcFlow2_Rate.mRun(mRun=>_cond[2])
	THEN;
		//
	ELSE;
		bCIP_Condition_Failed:=TRUE;
	END_IF	
END_IF

pcHeatExchanger.mRun_PID(Set_Point:=st_CIP_Param.r_Temper_DisInfection, controlManual:=g_Data.stHeatExchanger.bManual ,mRun_PID=>_temp);
tonr_CIP_Condition(PT:=SECOND_TO_TIME(tConditionTime));
IF TRUE 
AND pcHeatExchanger.mRun_With_SP(Set_Point:=st_CIP_Param.r_Temper_DisInfection, mRun_With_SP=>_cond[3])
//AND pcTemperature_Dis.mRun_With_SP(Set_Point:=st_CIP_Param.r_Temper_DisInfection, mRun_With_SP=>_cond[4])
AND pcTemp_ClntReturn.mRun_With_SP(Set_Point:=st_CIP_Param.r_Temper_DisInfection, mRun_With_SP=>_cond[5])
AND measure_Dis_2.x
AND TRUE
THEN;
	tonr_CIP_Condition.IN:=TRUE;
	m_MixProof_run();
ELSE;
	tonr_CIP_Condition.IN:=FALSE;
END_IF

IF NOT bSprinkler THEN;
	IF pcDisInfectant.mRun_With_SP(Set_Point:=st_CIP_Param.r_DisInfectionConcentration, mRun_With_SP=>_cond[6])
	AND tonr_CIP_Condition.IN
	THEN;
		//tonr_CIP_Condition.IN:=TRUE;
	ELSIF bSprinkler THEN;
		tonr_CIP_Condition.IN:=TRUE;
	ELSE;
		tonr_CIP_Condition.IN:=FALSE;
	END_IF	
END_IF	


IF tonr_CIP_Condition.Q 
AND bValveCleanDone
THEN
	bCIP_Condition_Done:=TRUE;
ELSE;
	bCIP_Condition_Done:=FALSE;	
END_IF


ton_Concentration_Filter(PT:=T#30S, IN:=stDisInfectant.Control_ON AND (NOT stDisInfectant.OverFlow) AND (NOT bSprinkler));
IF TRUE 	
AND ton_Concentration_Filter.Q	
THEN;
	bConcentration_correct:=TRUE;
ELSE;
	bConcentration_correct:=FALSE;
END_IF

// Reverce function
(*
IF Disinfct_Conc_Client_Done.x 
AND NOT pcDisInfectant.mRun()
AND NOT pcTemp_ClntReturn.mRun()
THEN;
	bCIP_Condition_Failed:=TRUE;
END_IF

IF Temperature_Dis_2_Done.x 
AND NOT pcTemperature_Dis.mRun()
THEN;
	bCIP_Condition_Failed:=TRUE;
END_IF


//ton_CIP_Condition(PT:=T#30S);
IF tConditionTime-nDisInf_CondActTime_Clnt>0 THEN
	tonr_CIP_Condition(PT:=SECOND_TO_TIME(tConditionTime-nDisInf_CondActTime_Clnt));
	bDisInf_CondActTime_Clnt_Done:=FALSE;
ELSE
	bDisInf_CondActTime_Clnt_Done:=TRUE;
END_IF
IF TRUE 
AND Disinfct_Conc_Client_Done.x
AND Temperature_Dis_2_Done.x
AND NOT bDisInf_CondActTime_Clnt_Done
AND TRUE
THEN;
	tonr_CIP_Condition.IN:=TRUE;
ELSE;
	nDisInf_CondActTime_Clnt:=TIME_TO_INT(tonr_CIP_Condition.ET)/1000;
	tonr_CIP_Condition.IN:=FALSE;
END_IF

IF tonr_CIP_Condition.Q 
OR bDisInf_CondActTime_Clnt_Done 
THEN;
	bCIP_Condition_Done:=TRUE;
ELSE;
	bCIP_Condition_Done:=FALSE;	
END_IF
*)
END_ACTION

ACTION _aCondition_CIP3_Client_exit:
tonr_CIP_Condition(IN:=FALSE);
END_ACTION

ACTION _aCondition_CIP3_Local_active:
fb_PumpCIP.m_Run(RPM:=pcFlow1_Rate.mRun_PID(Set_Point:=g_Data.arr_CIP_Param[E_CIP_Usage.eLocal].r_Flow_Pipe,controlManual:=NOT(fb_PumpCIP.modeAuto)));

IF TRUE 
AND pcFlow1_Rate.mRun(mRun=>_cond[1])
AND pcFlow2_Rate.mRun(mRun=>_cond[2])
//AND pcPressure.mRun()
THEN;
	//
ELSE;
	bCIP_Condition_Failed:=TRUE;
END_IF

pcHeatExchanger.mRun_PID(Set_Point:=g_Data.arr_CIP_Param[E_CIP_Usage.eLocal].r_Temper_DisInfection, controlManual:=g_Data.stHeatExchanger.bManual ,mRun_PID=>_temp);
tonr_CIP_Condition(PT:=SECOND_TO_TIME(g_Data.arr_CIP_Param[E_CIP_Usage.eLocal].t_ConditionDisInfection));
IF TRUE 
AND pcHeatExchanger.mRun_With_SP(Set_Point:=g_Data.arr_CIP_Param[E_CIP_Usage.eLocal].r_Temper_DisInfection, mRun_With_SP=>_cond[3])
AND pcTemperature_Dis.mRun_With_SP(Set_Point:=g_Data.arr_CIP_Param[E_CIP_Usage.eLocal].r_Temper_DisInfection, mRun_With_SP=>_cond[4])
AND pcTemp_ClntReturn.mRun_With_SP(Set_Point:=g_Data.arr_CIP_Param[E_CIP_Usage.eLocal].r_Temper_DisInfection, mRun_With_SP=>_cond[5])
AND pcDisInfectant.mRun_With_SP(Set_Point:=g_Data.arr_CIP_Param[E_CIP_Usage.eLocal].r_DisInfectionConcentration, mRun_With_SP=>_cond[6])	
AND measure_Dis.x
AND TRUE
THEN;
	tonr_CIP_Condition.IN:=TRUE;
ELSE;
	tonr_CIP_Condition.IN:=FALSE;
END_IF

IF tonr_CIP_Condition.Q THEN
	bCIP_Condition_Done:=TRUE;
ELSE;
	bCIP_Condition_Done:=FALSE;	
END_IF


ton_Concentration_Filter(PT:=T#30S, IN:=stDisInfectant.Control_ON AND NOT stDisInfectant.OverFlow);
IF TRUE 
AND ton_Concentration_Filter.Q	
THEN;
 bConcentration_correct:=TRUE;
ELSE;
 bConcentration_correct:=FALSE;
END_IF

// Reverce function
(*
IF Disinfct_Conc_Local_Done.x 
AND NOT pcDisInfectant.mRun()
THEN;
	bCIP_Condition_Failed:=TRUE;
END_IF

IF Temperature_Dis_1_Done.x 
AND NOT pcTemperature_Dis.mRun()
THEN;
	bCIP_Condition_Failed:=TRUE;
END_IF
*)
(*
//ton_CIP_Condition(PT:=T#30S);
IF g_Data.arr_CIP_Param[E_CIP_Usage.eLocal].t_ConditionDisInfection-nDisInf_CondActTime_Lcl>0 THEN
	tonr_CIP_Condition(PT:=SECOND_TO_TIME(g_Data.arr_CIP_Param[E_CIP_Usage.eLocal].t_ConditionDisInfection-nDisInf_CondActTime_Lcl));
	bDisInf_CondActTime_Lcl_Done:=FALSE;
ELSE
	bDisInf_CondActTime_Lcl_Done:=TRUE;
END_IF

IF TRUE 
AND Disinfct_Conc_Local_Done.x
AND Temperature_Dis_1_Done.x
AND NOT bDisInf_CondActTime_Lcl_Done
AND TRUE
THEN;
	tonr_CIP_Condition.IN:=TRUE;
ELSE;
	nDisInf_CondActTime_Lcl:=TIME_TO_INT(tonr_CIP_Condition.ET)/1000;
	tonr_CIP_Condition.IN:=FALSE;
END_IF

IF tonr_CIP_Condition.Q
OR bDisInf_CondActTime_Lcl_Done
THEN
	bCIP_Condition_Done:=TRUE;
ELSE;
	bCIP_Condition_Done:=FALSE;	
END_IF
*)
END_ACTION

ACTION _aCondition_CIP3_Local_exit:
tonr_CIP_Condition(IN:=FALSE);
END_ACTION

ACTION _aCondition_CIP4_Client_active:
IF NOT bSprinkler THEN
	//pipe
	tConditionTime	:=st_CIP_Param.t_ConditionWater;
	fFlowRate		:=st_CIP_Param.r_Flow_Pipe;
	
ELSE
	//sprinkler
	tConditionTime	:=st_CIP_Param.t_ConditionWater_Sprinkler;
	fFlowRate		:=st_CIP_Param.r_Flow_Sprinkler;
END_IF

IF Condition_CIP4_Client.t > SECOND_TO_TIME(st_CIP_Param.t_PumpInitRun) THEN;
	fb_PumpCIP.m_Run(RPM:=pcFlow1_Rate.mRun_PID(Set_Point:=fFlowRate,controlManual:=NOT(fb_PumpCIP.modeAuto)));
END_IF
fb_PumpClient.m_Run(RPM:=st_CIP_Param.r_CIP_Client_Pump);
//Level control

IF FALSE  
//AND (delta_T94_Volume < -st_CIP_Param.r_Volume_Recycle_Detergent AND eRefClient_fbElement.eState_Long=E_Element_State_Long.eCIP_2_Deterged
//OR delta_T94_Volume < -st_CIP_Param.r_Volume_Recycle_DisInfection AND eRefClient_fbElement.eState_Long=E_Element_State_Long.eCIP_4_Sanitized) 
OR lvlTank_T94.rTankLevel < 250
THEN;
	bCIP_Condition_Failed:=TRUE;
END_IF


// Connect return to R_Water
IF TRUE 
AND lvlTank_T93.rTankLevel<450 
AND fbCIP_Return.m_CheckStatus(eReqStatus:=E_CIP_Return.eDrain)
THEN;
	fbCIP_Return.m_Run(eReqProc:=E_CIP_Return.eT93_R_Water);
ELSE;
	
END_IF



// Connect return to Drain

IF TRUE 
AND lvlTank_T93.rTankLevel>500 // The tank is full
AND fbCIP_Return.m_CheckStatus(eReqStatus:=E_CIP_Return.eT93_R_Water)
THEN;
	fbCIP_Return.m_Run(eReqProc:=E_CIP_Return.eDrain);
ELSE;
	
END_IF

// Condition
tonr_CIP_Condition(PT:=SECOND_TO_TIME(tConditionTime));
IF bSprinkler THEN;
	IF TRUE 
	AND pcFlow1_Rate.mRun(mRun=>_cond[1])
	//AND pcFlow3_Rate.mRun(mRun=>_cond[2])
	THEN;
		tonr_CIP_Condition.IN:=TRUE;
	ELSE;
		tonr_CIP_Condition.IN:=FALSE;
	END_IF
ELSE;
	IF TRUE 
	AND pcFlow1_Rate.mRun(mRun=>_cond[1])
	//AND pcFlow2_Rate.mRun(mRun=>_cond[2])
	THEN;
		tonr_CIP_Condition.IN:=TRUE;
	ELSE;
		tonr_CIP_Condition.IN:=FALSE;
	END_IF	
	
END_IF

IF tonr_CIP_Condition.Q THEN
	bCIP_Condition_Done:=TRUE;
ELSE;
	bCIP_Condition_Done:=FALSE;	
END_IF

(*
IF TRUE 
AND bCIP_Condition_Done
OR bCIP_Condition_Failed
THEN;

ELSE;
	
END_IF

IF TRUE 
AND pcFlow1_Rate.mRun(mRun=>_cond[1])
AND pcFlow2_Rate.mRun(mRun=>_cond[2])
//AND pcPressure.mRun()
THEN;
	//
ELSE;
	bCIP_Condition_Failed:=TRUE;
END_IF
*)
END_ACTION

ACTION _aCondition_CIP4_Client_entry:
//fbCIP_Return.m_Run(eReqProc:=E_CIP_Return.eT93_R_Water);
bCIP_Condition_Failed:=FALSE;
bCIP_Condition_Done:=FALSE;
mVolumeReset_All();
END_ACTION

ACTION _aCondition_CIP4_Client_exit:
tonr_CIP_Condition(IN:=FALSE);
END_ACTION

ACTION _aConnect_CIP1_Drain_active:
bStepDone:=FALSE;

IF fbCIP_Source.m_CheckStatus(eReqStatus:=E_CIP_Source.eT93_R_Water) 
AND fbCIP_Usage.m_CheckStatus(eReqStatus:=eReq.eClient)
AND mCIP_Clients_status(command:=E_CIP_Client_Command.eCIP)
THEN

	CASE eReq.eClient OF	
		E_CIP_Usage.eTank_1:;
					bStepDone:=fbCIP_ClientTank_Marinade.m_CheckStatus(eReqStatus:=E_CIP_ClientTank.eTank_A);
					fbTank1.cip_Pump_linked:=TRUE;
		E_CIP_Usage.eTank_2:;
					bStepDone:=fbCIP_ClientTank_Marinade.m_CheckStatus(eReqStatus:=E_CIP_ClientTank.eTank_B);
					fbTank2.cip_Pump_linked:=TRUE;					
		E_CIP_Usage.eTank_3:;
					bStepDone:=fbCIP_ClientTank_Color.m_CheckStatus(eReqStatus:=E_CIP_ClientTank.eTank_A);
					fbTank3.cip_Pump_linked:=TRUE;					
		E_CIP_Usage.eTank_4:;
					bStepDone:=fbCIP_ClientTank_Color.m_CheckStatus(eReqStatus:=E_CIP_ClientTank.eTank_B);
					fbTank4.cip_Pump_linked:=TRUE;					
	ELSE;				
		bStepDone:=TRUE;
	END_CASE
	
END_IF
END_ACTION

ACTION _aConnect_CIP1_Drain_entry:
fbCIP_Source.m_Run(eReqProc:=E_CIP_Source.eT93_R_Water);
fbCIP_Usage.m_Run(eReqProc:=eReq.eClient);
mCIP_Clients_command(command:=E_CIP_Client_Command.eCIP);

CASE eReq.eClient OF

	E_CIP_Usage.eTank_1:;
				fbCIP_ClientTank_Marinade.m_Run(eReqProc:=E_CIP_ClientTank.eTank_A);
	E_CIP_Usage.eTank_2:;
				fbCIP_ClientTank_Marinade.m_Run(eReqProc:=E_CIP_ClientTank.eTank_B);	
	E_CIP_Usage.eTank_3:;
				fbCIP_ClientTank_Color.m_Run(eReqProc:=E_CIP_ClientTank.eTank_A);
	E_CIP_Usage.eTank_4:;
				fbCIP_ClientTank_Color.m_Run(eReqProc:=E_CIP_ClientTank.eTank_B);	

END_CASE

bSprinkler:=FALSE;

(*
CASE eReq.eClient OF
	E_CIP_Usage.eLocal:;
				//
	E_CIP_Usage.eTank_1:;
				fbCIP_ClientTank_Marinade.m_Run(eReqProc:=E_CIP_ClientTank.eTank_A);
	E_CIP_Usage.eTank_2:;
				fbCIP_ClientTank_Marinade.m_Run(eReqProc:=E_CIP_ClientTank.eTank_B);	
	E_CIP_Usage.eTank_3:;
				fbCIP_ClientTank_Color.m_Run(eReqProc:=E_CIP_ClientTank.eTank_A);
	E_CIP_Usage.eTank_4:;
				fbCIP_ClientTank_Color.m_Run(eReqProc:=E_CIP_ClientTank.eTank_A);	
	E_CIP_Usage.eTriBlender_Marinada,
	E_CIP_Usage.eLine_Marinada:;
				//
	E_CIP_Usage.eTriBlender_Color,
	E_CIP_Usage.eLine_Color:;
				//		
END_CASE
*)
END_ACTION

ACTION _aConnect_CIP2_01_active:
bStepDone:=FALSE;
IF fbCIP_Source.m_CheckStatus(eReqStatus:=E_CIP_Source.eT92_Detergent)  
AND fbCIP_Return.m_CheckStatus(eReqStatus:=E_CIP_Return.eT92_Detergent)  
AND fbPis.m_CheckByRecipe(stPis:=stPis_FillWater_T92, req:=E_Piston_Recipe_State.Release) THEN;
	bStepDone:=TRUE;
END_IF
END_ACTION

ACTION _aConnect_CIP2_01_entry:
fbCIP_Source.m_Run(eReqProc:=E_CIP_Source.eT92_Detergent);
fbCIP_Return.m_Run(eReqProc:=E_CIP_Return.eT92_Detergent);
fbPis.m_SetByRecipe(stPis:=stPis_FillWater_T92, req:=E_Piston_Recipe_State.Release);

m_DashState_done(stage:=E_CIP_DashStage_List.e03_CIP2_Local_Detergent_Fill);
m_DashState_activate(stage:=E_CIP_DashStage_List.e04_CIP2_Local_Detergent_Condition);
END_ACTION

ACTION _aConnect_CIP2_02_active:
bStepDone:=FALSE;
IF fbCIP_Return.m_CheckStatus(eReqStatus:=E_CIP_Return.eT92_Detergent)  
//AND fbPis.m_CheckByRecipe(stPis:=stPis_FillWater_T92, req:=E_Piston_Recipe_State.Release) 
THEN;
	bStepDone:=TRUE;
END_IF
END_ACTION

ACTION _aConnect_CIP2_02_entry:
fbCIP_Return.m_Run(eReqProc:=E_CIP_Return.eT92_Detergent);
fbPis.m_SetByRecipe(stPis:=stPis_FillWater_T92, req:=E_Piston_Recipe_State.Release);
//fb_PumpDetergent.m_Auto();
fb_HeatExchenger.m_Auto();

m_DashState_done(stage:=E_CIP_DashStage_List.e05_CIP2_Client_Detergent_Fill);
m_DashState_activate(stage:=E_CIP_DashStage_List.e06_CIP2_Client_Detergent_Condition_Pipe);
END_ACTION

ACTION _aConnect_CIP2_Drain_active:
bStepDone:=FALSE;
IF fbCIP_Usage.m_CheckStatus(eReqStatus:=eReq.eClient)  
AND fbCIP_Return.m_CheckStatus(eReqStatus:=E_CIP_Return.eDrain) 
AND mCIP_Clients_status(command:=E_CIP_Client_Command.eCIP)
THEN;

	CASE eReq.eClient OF	
		E_CIP_Usage.eTank_1:;
					bStepDone:=fbCIP_ClientTank_Marinade.m_CheckStatus(eReqStatus:=E_CIP_ClientTank.eTank_A);
					fbTank1.cip_Pump_linked:=TRUE;
		E_CIP_Usage.eTank_2:;
					bStepDone:=fbCIP_ClientTank_Marinade.m_CheckStatus(eReqStatus:=E_CIP_ClientTank.eTank_B);
					fbTank2.cip_Pump_linked:=TRUE;					
		E_CIP_Usage.eTank_3:;
					bStepDone:=fbCIP_ClientTank_Color.m_CheckStatus(eReqStatus:=E_CIP_ClientTank.eTank_A);
					fbTank3.cip_Pump_linked:=TRUE;					
		E_CIP_Usage.eTank_4:;
					bStepDone:=fbCIP_ClientTank_Color.m_CheckStatus(eReqStatus:=E_CIP_ClientTank.eTank_B);
					fbTank4.cip_Pump_linked:=TRUE;					
	ELSE;				
		bStepDone:=TRUE;
	END_CASE
	
END_IF

(*
	//eReq.eClient<>E_CIP_Usage.eLocal
	CASE eReq.eClient OF
		E_CIP_Usage.eTank_1:;
			//g_Data.fbTankTarget_1.m_Run(eReqProc:=E_Tank_Target.eCIP);
			IF g_Data.fbTankTarget_1.m_CheckStatus(eReqStatus:=E_Tank_Target.eCIP) THEN;
				bStepDone:=TRUE;
			ELSE;
				bStepDone:=FALSE;	
			END_IF
		E_CIP_Usage.eTank_2:;
			//g_Data.fbTankTarget_2.m_Run(eReqProc:=E_Tank_Target.eCIP);
			IF g_Data.fbTankTarget_2.m_CheckStatus(eReqStatus:=E_Tank_Target.eCIP) THEN;
				bStepDone:=TRUE;
			ELSE;
				bStepDone:=FALSE;	
			END_IF	
		E_CIP_Usage.eTank_3:;
			//g_Data.fbTankTarget_3.m_Run(eReqProc:=E_Tank_Target.eCIP);
			IF g_Data.fbTankTarget_3.m_CheckStatus(eReqStatus:=E_Tank_Target.eCIP) THEN;
				bStepDone:=TRUE;
			ELSE;
				bStepDone:=FALSE;	
			END_IF	
		E_CIP_Usage.eTank_4:;
			//g_Data.fbTankTarget_4.m_Run(eReqProc:=E_Tank_Target.eCIP);
			IF g_Data.fbTankTarget_4.m_CheckStatus(eReqStatus:=E_Tank_Target.eCIP) THEN;
				bStepDone:=TRUE;
			ELSE;
				bStepDone:=FALSE;	
			END_IF	
		E_CIP_Usage.eTriBlender_Marinada:;
			//g_Data.fbTriBlenderSource_Marinade.m_Run(eReqProc:=E_Line_Source.eCIP);	
			//g_Data.fbTriBlenderTarget_Marinade.m_Run(eReqProc:=E_Line_Target.eCIP);	
			IF  g_Data.fbTriBlenderSource_Marinade.m_CheckStatus(eReqStatus:=E_Line_Source.eCIP) 
			AND g_Data.fbTriBlenderTarget_Marinade.m_CheckStatus(eReqStatus:=E_Line_Target.eCIP) THEN;
				bStepDone:=TRUE;
			ELSE;
				bStepDone:=FALSE;	
			END_IF
		E_CIP_Usage.eTriBlender_Color:;
			//g_Data.fbTriBlenderSource_Color.m_Run(eReqProc:=E_Line_Source.eCIP);	
			//g_Data.fbTriBlenderTarget_Color.m_Run(eReqProc:=E_Line_Target.eCIP);
			IF  g_Data.fbTriBlenderSource_Color.m_CheckStatus(eReqStatus:=E_Line_Source.eCIP) 
			AND g_Data.fbTriBlenderTarget_Color.m_CheckStatus(eReqStatus:=E_Line_Target.eCIP) THEN;
				bStepDone:=TRUE;
			ELSE;
				bStepDone:=FALSE;	
			END_IF		
		E_CIP_Usage.eLine_Marinada:;
			//g_Data.fbLineSource_Marinade.m_Run(eReqProc:=E_Line_Source.eCIP);	
			//g_Data.fbLineTarget_Marinade.m_Run(eReqProc:=E_Line_Target.eCIP);
			IF  g_Data.fbLineSource_Marinade.m_CheckStatus(eReqStatus:=E_Line_Source.eCIP) 
			AND g_Data.fbLineTarget_Marinade.m_CheckStatus(eReqStatus:=E_Line_Target.eCIP) THEN;
				bStepDone:=TRUE;
			ELSE;
				bStepDone:=FALSE;	
			END_IF	
		E_CIP_Usage.eLine_Color:;
			//g_Data.fbLineSource_Color.m_Run(eReqProc:=E_Line_Source.eCIP);	
			//g_Data.fbLineTarget_Color.m_Run(eReqProc:=E_Line_Target.eCIP);
			IF  g_Data.fbLineSource_Color.m_CheckStatus(eReqStatus:=E_Line_Source.eCIP) 
			AND g_Data.fbLineTarget_Color.m_CheckStatus(eReqStatus:=E_Line_Target.eCIP) THEN;
				bStepDone:=TRUE;
			ELSE;
				bStepDone:=FALSE;	
			END_IF	
	ELSE;
		//wrong, - local
		bStepDone:=FALSE;
	END_CASE
*)
END_ACTION

ACTION _aConnect_CIP2_Drain_entry:
fbCIP_Usage.m_Run(eReqProc:=eReq.eClient);
fbCIP_Return.m_Run(eReqProc:=E_CIP_Return.eDrain);
fb_HeatExchenger.m_Auto();

mCIP_Clients_command(command:=E_CIP_Client_Command.eCIP);

CASE eReq.eClient OF

	E_CIP_Usage.eTank_1:;
				fbCIP_ClientTank_Marinade.m_Run(eReqProc:=E_CIP_ClientTank.eTank_A);
	E_CIP_Usage.eTank_2:;
				fbCIP_ClientTank_Marinade.m_Run(eReqProc:=E_CIP_ClientTank.eTank_B);	
	E_CIP_Usage.eTank_3:;
				fbCIP_ClientTank_Color.m_Run(eReqProc:=E_CIP_ClientTank.eTank_A);
	E_CIP_Usage.eTank_4:;
				fbCIP_ClientTank_Color.m_Run(eReqProc:=E_CIP_ClientTank.eTank_B);	

END_CASE

m_DashState_activate(stage:=E_CIP_DashStage_List.e05_CIP2_Client_Detergent_Fill);
END_ACTION

ACTION _aConnect_CIP3_01_active:
bStepDone:=FALSE;
IF fbCIP_Source.m_CheckStatus(eReqStatus:=E_CIP_Source.eT91_Sanitation)  
AND fbCIP_Return.m_CheckStatus(eReqStatus:=E_CIP_Return.eT91_Sanitation)  
AND fbPis.m_CheckByRecipe(stPis:=stPis_FillWater_T91, req:=E_Piston_Recipe_State.Release) THEN;
	bStepDone:=TRUE;
END_IF
END_ACTION

ACTION _aConnect_CIP3_01_entry:
fbCIP_Source.m_Run(eReqProc:=E_CIP_Source.eT91_Sanitation);
fbCIP_Return.m_Run(eReqProc:=E_CIP_Return.eT91_Sanitation);
fbPis.m_SetByRecipe(stPis:=stPis_FillWater_T91, req:=E_Piston_Recipe_State.Release);
tonr_CIP_Condition(ResetTime:=TRUE);

m_DashState_done(stage:=E_CIP_DashStage_List.e12_CIP4_Local_DisInfection_Fill);
m_DashState_activate(stage:=E_CIP_DashStage_List.e13_CIP4_Local_DisInfection_Condition);
END_ACTION

ACTION _aConnect_CIP3_02_active:
bStepDone:=FALSE;
IF fbCIP_Return.m_CheckStatus(eReqStatus:=E_CIP_Return.eT91_Sanitation)  
//AND fbPis.m_CheckByRecipe(stPis:=stPis_FillWater_T92, req:=E_Piston_Recipe_State.Release) 
THEN;
	bStepDone:=TRUE;
END_IF
END_ACTION

ACTION _aConnect_CIP3_02_entry:
fbCIP_Return.m_Run(eReqProc:=E_CIP_Return.eT91_Sanitation);

m_DashState_done(stage:=E_CIP_DashStage_List.e14_CIP4_Client_DisInfection_Fill);
m_DashState_activate(stage:=E_CIP_DashStage_List.e15_CIP4_Client_DisInfection_Condition_Pipe);
END_ACTION

ACTION _aConnect_CIP3_Drain_active:
bStepDone:=FALSE;
IF fbCIP_Usage.m_CheckStatus(eReqStatus:=eReq.eClient)  
AND fbCIP_Return.m_CheckStatus(eReqStatus:=E_CIP_Return.eDrain) 
AND mCIP_Clients_status(command:=E_CIP_Client_Command.eCIP)
THEN;

	CASE eReq.eClient OF	
		E_CIP_Usage.eTank_1:;
					bStepDone:=fbCIP_ClientTank_Marinade.m_CheckStatus(eReqStatus:=E_CIP_ClientTank.eTank_A);
					fbTank1.cip_Pump_linked:=TRUE;
		E_CIP_Usage.eTank_2:;
					bStepDone:=fbCIP_ClientTank_Marinade.m_CheckStatus(eReqStatus:=E_CIP_ClientTank.eTank_B);
					fbTank2.cip_Pump_linked:=TRUE;					
		E_CIP_Usage.eTank_3:;
					bStepDone:=fbCIP_ClientTank_Color.m_CheckStatus(eReqStatus:=E_CIP_ClientTank.eTank_A);
					fbTank3.cip_Pump_linked:=TRUE;					
		E_CIP_Usage.eTank_4:;
					bStepDone:=fbCIP_ClientTank_Color.m_CheckStatus(eReqStatus:=E_CIP_ClientTank.eTank_B);
					fbTank4.cip_Pump_linked:=TRUE;					
	ELSE;				
		bStepDone:=TRUE;
	END_CASE
	
END_IF
END_ACTION

ACTION _aConnect_CIP3_Drain_entry:
fbCIP_Usage.m_Run(eReqProc:=eReq.eClient);
fbCIP_Return.m_Run(eReqProc:=E_CIP_Return.eDrain);
fb_HeatExchenger.m_Auto();

mCIP_Clients_command(command:=E_CIP_Client_Command.eCIP);

CASE eReq.eClient OF

	E_CIP_Usage.eTank_1:;
				fbCIP_ClientTank_Marinade.m_Run(eReqProc:=E_CIP_ClientTank.eTank_A);
	E_CIP_Usage.eTank_2:;
				fbCIP_ClientTank_Marinade.m_Run(eReqProc:=E_CIP_ClientTank.eTank_B);	
	E_CIP_Usage.eTank_3:;
				fbCIP_ClientTank_Color.m_Run(eReqProc:=E_CIP_ClientTank.eTank_A);
	E_CIP_Usage.eTank_4:;
				fbCIP_ClientTank_Color.m_Run(eReqProc:=E_CIP_ClientTank.eTank_B);	

END_CASE

m_DashState_activate(stage:=E_CIP_DashStage_List.e14_CIP4_Client_DisInfection_Fill);
END_ACTION

ACTION _aConnect_CIP4_active:
bStepDone:=FALSE;
IF TRUE
AND fbCIP_Source.m_CheckStatus(eReqStatus:=E_CIP_Source.eT94_Water) 
//AND fbCIP_Source.m_CheckStatus(eReqStatus:=E_CIP_Source.eT93_R_Water) 
AND fbCIP_Usage.m_CheckStatus(eReqStatus:=eReq.eClient)  
//AND fbCIP_Return.m_CheckStatus(eReqStatus:=E_CIP_Return.eDrain) 
AND mCIP_Clients_status(command:=E_CIP_Client_Command.eCIP)
THEN;

	CASE eReq.eClient OF	
		E_CIP_Usage.eTank_1:;
					bStepDone:=fbCIP_ClientTank_Marinade.m_CheckStatus(eReqStatus:=E_CIP_ClientTank.eTank_A);
					fbTank1.cip_Pump_linked:=TRUE;
		E_CIP_Usage.eTank_2:;
					bStepDone:=fbCIP_ClientTank_Marinade.m_CheckStatus(eReqStatus:=E_CIP_ClientTank.eTank_B);
					fbTank2.cip_Pump_linked:=TRUE;					
		E_CIP_Usage.eTank_3:;
					bStepDone:=fbCIP_ClientTank_Color.m_CheckStatus(eReqStatus:=E_CIP_ClientTank.eTank_A);
					fbTank3.cip_Pump_linked:=TRUE;					
		E_CIP_Usage.eTank_4:;
					bStepDone:=fbCIP_ClientTank_Color.m_CheckStatus(eReqStatus:=E_CIP_ClientTank.eTank_B);
					fbTank4.cip_Pump_linked:=TRUE;					
	ELSE;				
		bStepDone:=TRUE;
	END_CASE
	
END_IF

IF bStepDone THEN;
	CASE eRefClient_fbElement.eState_Long OF
		E_Element_State_Long.eCIP_2_Deterged:;
				//fbCIP_Return.m_Run(eReqProc:=E_CIP_Return.eT92_Detergent);
				bStepDone:=fbCIP_Return.m_CheckStatus(eReqStatus:=E_CIP_Return.eT92_Detergent);
		E_Element_State_Long.eCIP_4_Sanitized:;
				//fbCIP_Return.m_Run(eReqProc:=E_CIP_Return.eT91_Sanitation);	
				bStepDone:=fbCIP_Return.m_CheckStatus(eReqStatus:=E_CIP_Return.eT91_Sanitation);
	ELSE;
		bStepDone:=FALSE;
	END_CASE	
END_IF
END_ACTION

ACTION _aConnect_CIP4_entry:
fbCIP_Source.m_Run(eReqProc:=E_CIP_Source.eT94_Water);
//Temp solution for T93
//fbCIP_Source.m_Run(eReqProc:=E_CIP_Source.eT93_R_Water);
fbCIP_Usage.m_Run(eReqProc:=eReq.eClient);

mCIP_Clients_command(command:=E_CIP_Client_Command.eCIP);



CASE eRefClient_fbElement.eState_Long OF
	E_Element_State_Long.eCIP_2_Deterged:;
			fbCIP_Return.m_Run(eReqProc:=E_CIP_Return.eT92_Detergent);
		
	E_Element_State_Long.eCIP_4_Sanitized:;
			fbCIP_Return.m_Run(eReqProc:=E_CIP_Return.eT91_Sanitation);				
END_CASE

CASE eReq.eClient OF

	E_CIP_Usage.eTank_1:;
				fbCIP_ClientTank_Marinade.m_Run(eReqProc:=E_CIP_ClientTank.eTank_A);
	E_CIP_Usage.eTank_2:;
				fbCIP_ClientTank_Marinade.m_Run(eReqProc:=E_CIP_ClientTank.eTank_B);	
	E_CIP_Usage.eTank_3:;
				fbCIP_ClientTank_Color.m_Run(eReqProc:=E_CIP_ClientTank.eTank_A);
	E_CIP_Usage.eTank_4:;
				fbCIP_ClientTank_Color.m_Run(eReqProc:=E_CIP_ClientTank.eTank_B);	

END_CASE
END_ACTION

ACTION _aConnect_CIP4_R_Water_active:
bStepDone:=FALSE;
IF fbCIP_Return.m_CheckStatus(eReqStatus:=E_CIP_Return.eT93_R_Water)  
THEN;
	bStepDone:=TRUE;
END_IF
END_ACTION

ACTION _aConnect_CIP4_R_Water_entry:
fbCIP_Return.m_Run(eReqProc:=E_CIP_Return.eT93_R_Water);
mVolumeReset_All();

	CASE eRefClient_fbElement.eState_Long OF
	
		E_Element_State_Long.eCIP_2_Deterged:;
				m_DashState_done(stage:=E_CIP_DashStage_List.e09_CIP3_Detergent_Drain);
				m_DashState_activate(stage:=E_CIP_DashStage_List.e10_CIP3_Detergent_Clean_Pipe);
	
		E_Element_State_Long.eCIP_4_Sanitized:;
				m_DashState_done(stage:=E_CIP_DashStage_List.e18_CIP5_DisInfection_Drain);
				m_DashState_activate(stage:=E_CIP_DashStage_List.e19_CIP5_DisInfection_Clean_Pipe);
				
	END_CASE
END_ACTION

ACTION _aDeterg_Dose_1_active:

bStepDone:=fb_PumpDetergent.m_RunVolume(Volume:=0.9*(lvlTank_T92.rTankLevel*stDetergent.Deviation*10)); // 10= 1Litr*1000cc/100%
END_ACTION

ACTION _aDeterg_Dose_2_active:

bStepDone:=fb_PumpDetergent.m_RunVolume(Volume:=0.9*(lvlTank_T92.rTankLevel*stDetergent.Deviation*10)); // 10= 1Litr*1000cc/100%
END_ACTION

ACTION _aDeterg_Overflow_1_active:
IF lvlTank_T92.rTankLevel>=rDeluteVolume OR bCIP_Condition_Failed  THEN;	
	bStepDone:=TRUE;
	fbPis.m_SetByRecipe(stPis:=stPis_FillWater_T92, req:=E_Piston_Recipe_State.Release);
ELSE;
	//Fill water
	bStepDone:=FALSE;
	IF NOT arrTanksSens[E_Tank_Name.T92].get_stTankLevel_OverFlow() THEN;
		fbPis.m_SetByRecipe(stPis:=stPis_FillWater_T92, req:=E_Piston_Recipe_State.Act);			
	END_IF	
END_IF
END_ACTION

ACTION _aDeterg_Overflow_1_entry:
rDeltaWater_DeterLocal:=m_OverFlowCorrect(
							rTc:=stDetergent.rSetPoint , //g_Data.arr_CIP_Param[E_CIP_Usage.eLocal].r_DetergentConcentration
							rAv:=lvlTank_T92.rTankLevel , 
							rAc:=stDetergent.rValue );

fbPrintErrMessageByID(sModuleDescription:='CIP',sActErrorID:='101x000x101');							
rDeluteVolume:=rDeltaWater_DeterLocal + lvlTank_T92.rTankLevel;

IF rDeluteVolume>rDeluteVolume_max THEN;
	// message
	iConcentrationDeluteCounter:=iConcentrationDeluteCounter+1;
	IF iConcentrationDeluteCounter>3 THEN;
		fbPrintErrMessageByID(sModuleDescription:='eCIP',sActErrorID:='101x000x103');
	ELSE;
		fbPrintErrMessageByID(sModuleDescription:='CIP',sActErrorID:='101x000x102');
	END_IF
	rDeluteVolume:=rDeluteVolume_max;
END_IF
END_ACTION

ACTION _aDeterg_Overflow_2_active:
IF lvlTank_T92.rTankLevel>=rDeluteVolume OR bCIP_Condition_Failed THEN;	
	bStepDone:=TRUE;
	fbPis.m_SetByRecipe(stPis:=stPis_FillWater_T92, req:=E_Piston_Recipe_State.Release);
ELSE;
	//Fill water
	bStepDone:=FALSE;
	IF NOT arrTanksSens[E_Tank_Name.T92].get_stTankLevel_OverFlow() THEN;
		fbPis.m_SetByRecipe(stPis:=stPis_FillWater_T92, req:=E_Piston_Recipe_State.Act);			
	END_IF	
END_IF
END_ACTION

ACTION _aDeterg_Overflow_2_entry:
rDeltaWater_DeterClient:=m_OverFlowCorrect(
							rTc:=stDetergent.rSetPoint , 
							rAv:=lvlTank_T92.rTankLevel , 
							rAc:=stDetergent.rValue );
							
fbPrintErrMessageByID(sModuleDescription:='CIP',sActErrorID:='101x000x101');							
rDeluteVolume:=rDeltaWater_DeterClient + lvlTank_T92.rTankLevel;

IF rDeluteVolume>rDeluteVolume_max THEN;
	// message
	iConcentrationDeluteCounter:=iConcentrationDeluteCounter+1;
	IF iConcentrationDeluteCounter>3 THEN;
		fbPrintErrMessageByID(sModuleDescription:='eCIP',sActErrorID:='101x000x103');
	ELSE;
		fbPrintErrMessageByID(sModuleDescription:='CIP',sActErrorID:='101x000x102');
	END_IF
	rDeluteVolume:=rDeluteVolume_max;
END_IF
END_ACTION

ACTION _aDisconnect_n_Drain_CIP_Client_active:
bStepDone:=FALSE;

IF fbCIP_Source.m_CheckStatus(eReqStatus:=E_CIP_Source.eClose) 
AND fbCIP_Usage.m_CheckStatus(eReqStatus:=E_CIP_Usage.eLocal) 
AND fbCIP_Return.m_CheckStatus(eReqStatus:=E_CIP_Return.eDrain)
AND mCIP_Clients_status(command:=E_CIP_Client_Command.eClose)
THEN

	CASE eReq.eClient OF
	
		E_CIP_Usage.eTank_1:;
					bStepDone:=fbCIP_ClientTank_Marinade.m_CheckStatus(eReqStatus:=E_CIP_ClientTank.eClose);
		E_CIP_Usage.eTank_2:;
					bStepDone:=fbCIP_ClientTank_Marinade.m_CheckStatus(eReqStatus:=E_CIP_ClientTank.eClose);	
		E_CIP_Usage.eTank_3:;
					bStepDone:=fbCIP_ClientTank_Color.m_CheckStatus(eReqStatus:=E_CIP_ClientTank.eClose);
		E_CIP_Usage.eTank_4:;
					bStepDone:=fbCIP_ClientTank_Color.m_CheckStatus(eReqStatus:=E_CIP_ClientTank.eClose);	
		E_CIP_Usage.eTriBlender_Color,
		E_CIP_Usage.eTriBlender_Marinada:;
					bStepDone:=fbTriBlender_Select.m_CheckStatus(eReqStatus:=E_TriBlenderSelect.eMarinade);											
	ELSE;				
		bStepDone:=TRUE;
	END_CASE
	
END_IF

fbTank1.cip_Pump_linked:=FALSE;
fbTank2.cip_Pump_linked:=FALSE;
fbTank3.cip_Pump_linked:=FALSE;
fbTank4.cip_Pump_linked:=FALSE;

(* old, before drain done validation
IF fbCIP_Source.m_CheckStatus(eReqStatus:=E_CIP_Source.eClose) 
AND fbCIP_Usage.m_CheckStatus(eReqStatus:=E_CIP_Usage.eLocal) 
AND fbCIP_Return.m_CheckStatus(eReqStatus:=E_CIP_Return.eDrain)
AND mCIP_Clients_status(command:=E_CIP_Client_Command.eDrain)
THEN

	CASE eReq.eClient OF
	
		E_CIP_Usage.eTank_1:;
					bStepDone:=fbCIP_ClientTank_Marinade.m_CheckStatus(eReqStatus:=E_CIP_ClientTank.eDrain);
		E_CIP_Usage.eTank_2:;
					bStepDone:=fbCIP_ClientTank_Marinade.m_CheckStatus(eReqStatus:=E_CIP_ClientTank.eDrain);	
		E_CIP_Usage.eTank_3:;
					bStepDone:=fbCIP_ClientTank_Color.m_CheckStatus(eReqStatus:=E_CIP_ClientTank.eDrain);
		E_CIP_Usage.eTank_4:;
					bStepDone:=fbCIP_ClientTank_Color.m_CheckStatus(eReqStatus:=E_CIP_ClientTank.eDrain);	
		E_CIP_Usage.eTriBlender_Color,
		E_CIP_Usage.eTriBlender_Marinada:;
					bStepDone:=fbTriBlender_Select.m_CheckStatus(eReqStatus:=E_TriBlenderSelect.eDrain);											
	ELSE;				
		bStepDone:=TRUE;
	END_CASE
	
END_IF
*)
END_ACTION

ACTION _aDisconnect_n_Drain_CIP_Client_entry:
fbCIP_Source.m_Run(eReqProc:=E_CIP_Source.eClose);
fbCIP_Usage.m_Run(eReqProc:=E_CIP_Usage.eLocal);
fbCIP_Return.m_Run(eReqProc:=E_CIP_Return.eDrain);
mCIP_Clients_command(command:=E_CIP_Client_Command.eDrain);

IF bClientTypeIs_Tank THEN;
	fb_Stirrer.m_Stop();
END_IF

CASE eReq.eClient OF

	E_CIP_Usage.eTank_1:;
				fbCIP_ClientTank_Marinade.m_Run(eReqProc:=E_CIP_ClientTank.eDrain);
	E_CIP_Usage.eTank_2:;
				fbCIP_ClientTank_Marinade.m_Run(eReqProc:=E_CIP_ClientTank.eDrain);	
	E_CIP_Usage.eTank_3:;
				fbCIP_ClientTank_Color.m_Run(eReqProc:=E_CIP_ClientTank.eDrain);
	E_CIP_Usage.eTank_4:;
				fbCIP_ClientTank_Color.m_Run(eReqProc:=E_CIP_ClientTank.eDrain);	

END_CASE

IF __ISVALIDREF(eRefClient_fbElement) THEN;
	IF eRefClient_fbElement.eElementID=E_Element_List.eTriBlender_Marinada THEN;
		fbTriBlender_Select.m_Run(eReqProc:=E_TriBlenderSelect.eDrain);
	END_IF
	
	IF eRefClient_fbElement.eElementID=E_Element_List.eTriBlender_Color THEN;
		fbTriBlender_Select.m_Run(eReqProc:=E_TriBlenderSelect.eDrain);
	END_IF	
END_IF
END_ACTION

ACTION _aDisconnect_Old_Client_entry:
eReq:=eReqBlank;
eRun:=E_CIP_Source.eNone;
m_CleanEmpty_Spaces();

IF __ISVALIDREF(eRefClient_fbElement) THEN;
	IF eRefClient_fbElement.m_Get_CIP_Avilable() THEN;
		eRefClient_fbElement.m_Disconnect();
	END_IF
END_IF
eRefClient_fbElement REF= fbElement_Blank;

m_Disconnect_All_Client();
m_DashState_MixProof_set();
END_ACTION

ACTION _aDisinfct_Dose_1_active:

bStepDone:=fb_PumpDisinfection.m_RunVolume(Volume:=0.9*(lvlTank_T91.rTankLevel*stDisInfectant.Deviation*10)); // 10= 1Litr*1000cc/100%
END_ACTION

ACTION _aDisinfct_Dose_2_active:

bStepDone:=fb_PumpDisinfection.m_RunVolume(Volume:=0.9*(lvlTank_T91.rTankLevel*stDisInfectant.Deviation*10)); // 10= 1Litr*1000cc/100%
END_ACTION

ACTION _aDisinfct_Overflow_1_active:
IF lvlTank_T91.rTankLevel>=rDeluteVolume OR bCIP_Condition_Failed  THEN;	
	bStepDone:=TRUE;
	fbPis.m_SetByRecipe(stPis:=stPis_FillWater_T91, req:=E_Piston_Recipe_State.Release);
ELSE;
	//Fill water
	bStepDone:=FALSE;
	IF NOT arrTanksSens[E_Tank_Name.T91].get_stTankLevel_OverFlow() THEN;
		fbPis.m_SetByRecipe(stPis:=stPis_FillWater_T91, req:=E_Piston_Recipe_State.Act);			
	END_IF	
END_IF
END_ACTION

ACTION _aDisinfct_Overflow_1_entry:
rDeltaWater_DisInfLocal:=m_OverFlowCorrect(
								rTc:=stDisInfectant.rSetPoint , //g_Data.arr_CIP_Param[E_CIP_Usage.eLocal].r_DisInfectionConcentration
								rAv:=lvlTank_T91.rTankLevel , 
								rAc:=stDisInfectant.rValue );
								
fbPrintErrMessageByID(sModuleDescription:='CIP',sActErrorID:='101x000x111');							
rDeluteVolume:=rDeltaWater_DisInfLocal + lvlTank_T91.rTankLevel;

IF rDeluteVolume>rDeluteVolume_max THEN;
	// message
	iConcentrationDeluteCounter:=iConcentrationDeluteCounter+1;
	IF iConcentrationDeluteCounter>3 THEN;
		fbPrintErrMessageByID(sModuleDescription:='eCIP',sActErrorID:='101x000x113');
	ELSE;
		fbPrintErrMessageByID(sModuleDescription:='CIP',sActErrorID:='101x000x112');
	END_IF
	
	rDeluteVolume:=rDeluteVolume_max;
END_IF
END_ACTION

ACTION _aDisinfct_Overflow_2_active:
IF lvlTank_T91.rTankLevel>=rDeluteVolume OR bCIP_Condition_Failed  THEN;	
	bStepDone:=TRUE;
	fbPis.m_SetByRecipe(stPis:=stPis_FillWater_T91, req:=E_Piston_Recipe_State.Release);
ELSE;
	//Fill water
	bStepDone:=FALSE;
	IF NOT arrTanksSens[E_Tank_Name.T91].get_stTankLevel_OverFlow() THEN;
		fbPis.m_SetByRecipe(stPis:=stPis_FillWater_T91, req:=E_Piston_Recipe_State.Act);			
	END_IF	
END_IF
END_ACTION

ACTION _aDisinfct_Overflow_2_entry:
rDeltaWater_DisInfClient:=m_OverFlowCorrect(
								rTc:=stDisInfectant.rSetPoint , 
								rAv:=lvlTank_T91.rTankLevel , 
								rAc:=stDisInfectant.rValue );
								
fbPrintErrMessageByID(sModuleDescription:='CIP',sActErrorID:='101x000x111');							
rDeluteVolume:=rDeltaWater_DisInfClient + lvlTank_T91.rTankLevel;

IF rDeluteVolume>rDeluteVolume_max THEN;
	// message
	iConcentrationDeluteCounter:=iConcentrationDeluteCounter+1;
	IF iConcentrationDeluteCounter>3 THEN;
		fbPrintErrMessageByID(sModuleDescription:='eCIP',sActErrorID:='101x000x113');
	ELSE;
		fbPrintErrMessageByID(sModuleDescription:='CIP',sActErrorID:='101x000x112');
	END_IF
	
	rDeluteVolume:=rDeluteVolume_max;
END_IF
END_ACTION

ACTION _aDone_entry:
eRefClient_fbElement.m_Disconnect();
arCIP_RequestBufer[0]:=eReqBlank;
bRun:=FALSE;
END_ACTION

ACTION _aEnd_Check_active:
bStepDone:=FALSE;
IF TRUE 
AND eRefClient_fbElement.eState_Long = E_Element_State_Long.eCIP_1_Rinzed
AND eReq.eType = E_CIP_Type.R_Water
AND eReq.eClient<>E_CIP_Usage.eLocal
THEN;
	bStepDone:=TRUE;
	
ELSIF TRUE 
AND eRefClient_fbElement.eState_Long = E_Element_State_Long.eCIP_3_Deterged_Clean
AND eReq.eType = E_CIP_Type.Detergent
//AND eReq.eClient=E_CIP_Usage.eLocal
THEN;
	bStepDone:=TRUE;
	
ELSIF TRUE 
AND eRefClient_fbElement.eState_Long = E_Element_State_Long.eCIP_5_Done
AND eReq.eType = E_CIP_Type.Full
//AND eReq.eClient<>E_CIP_Usage.eLocal
THEN;
	bStepDone:=TRUE;
	
END_IF
END_ACTION

ACTION _aFill_For_MixProof_CIP2_active:
bStepDone:=m_ClientTank_Level_IsHigher_Then(min_Level:=50);
END_ACTION

ACTION _aFill_For_MixProof_CIP2_entry:
bSprinkler:=TRUE;
fb_PumpCIP.m_Run(RPM:=st_CIP_Param.r_CIP_Pump);
fb_PumpClient.m_Stop();

m_MixProof_set();
END_ACTION

ACTION _aFill_For_MixProof_CIP3_active:
bStepDone:=m_ClientTank_Level_IsHigher_Then(min_Level:=50);
END_ACTION

ACTION _aFill_For_MixProof_CIP3_entry:
bSprinkler:=TRUE;
fb_PumpCIP.m_Run(RPM:=st_CIP_Param.r_CIP_Pump);
fb_PumpClient.m_Stop();

m_MixProof_set();
END_ACTION

ACTION _aFill_Solution_CIP2_active:
bStepDone:=FALSE;
volume_Requered:= REAL_TO_INT(st_CIP_Param.r_Volume_Solution_Fill);
volume_Actual:= REAL_TO_INT(-delta_T92_Volume);

IF volume_Actual >= volume_Requered THEN;
	bStepDone:=TRUE;
END_IF
END_ACTION

ACTION _aFill_Solution_CIP3_active:
fb_PumpCIP.m_Run(RPM:=st_CIP_Param.r_CIP_Pump);
fb_PumpClient.m_Run(RPM:=st_CIP_Param.r_CIP_Client_Pump);

bStepDone:=FALSE;
volume_Requered:= REAL_TO_INT(st_CIP_Param.r_Volume_Solution_Fill);
volume_Actual:= REAL_TO_INT(-delta_T91_Volume);

IF volume_Actual >= volume_Requered THEN;
	bStepDone:=TRUE;
END_IF
END_ACTION

ACTION _aFill_Solution_CIP3_entry:
mVolumeReset_All();
tonr_CIP_Condition(ResetTime:=TRUE);
END_ACTION

ACTION _aFill_Water_T91_active:
nDisInf_CondActTime_Lcl:=0;
nDisInf_CondActTime_Clnt:=0;
bDisInf_CondActTime_Lcl_Done:=FALSE;
bDisInf_CondActTime_Clnt_Done:=FALSE;

bStepDone:=FALSE;
IF fbCIP_Source.m_CheckStatus(eReqStatus:=E_CIP_Source.eClose) 
AND fbCIP_Usage.m_CheckStatus(eReqStatus:=E_CIP_Usage.eLocal)  
AND fbCIP_Return.m_CheckStatus(eReqStatus:=E_CIP_Return.eDrain)  
//AND fbPis.m_CheckByRecipe(stPis:=stPis_FillWater_T91, req:=E_Piston_Recipe_State.Act) 
THEN;
	//IF eReq.eClient=E_CIP_Usage.eLocal 
	IF lvlTank_T91.e_state=E_Tank_Level.eLL
	AND lvlTank_T91.rTankLevel>g_Data.arr_CIP_Param[E_CIP_Usage.eLocal].r_Tank91_Volume//250 // Local requered Level
	THEN;	
		bStepDone:=TRUE;
		fbPis.m_SetByRecipe(stPis:=stPis_FillWater_T91, req:=E_Piston_Recipe_State.Release);
	(*ELSIF lvlTank_T91.e_state=E_Tank_Level.eLL
	AND lvlTank_T91.rTankLevel>g_Data.arr_CIP_Param[E_CIP_Usage.eLocal].r_TankLevel_2//300 // Client requered Level
	THEN;
		//Level OK
		bStepDone:=TRUE;
		fbPis.m_SetByRecipe(stPis:=stPis_FillWater_T91, req:=E_Piston_Recipe_State.Release);*)
	ELSE;
		//Fill water
		IF NOT arrTanksSens[E_Tank_Name.T91].get_stTankLevel_OverFlow() THEN;
			fbPis.m_SetByRecipe(stPis:=stPis_FillWater_T91, req:=E_Piston_Recipe_State.Act);			
		END_IF	
	END_IF	
END_IF
END_ACTION

ACTION _aFill_Water_T91_entry:
fbCIP_Source.m_Run(eReqProc:=E_CIP_Source.eClose);
fbCIP_Usage.m_Run(eReqProc:=E_CIP_Usage.eLocal);
fbCIP_Return.m_Run(eReqProc:=E_CIP_Return.eDrain);
bSprinkler:=FALSE;

m_DashState_activate(stage:=E_CIP_DashStage_List.e12_CIP4_Local_DisInfection_Fill);
	
m_MixProof_set();
END_ACTION

ACTION _aFill_Water_T92_active:
//Reset
nDeter_CondActTime_Lcl:=0;
nDeter_CondActTime_Clnt:=0;
bDeter_CondActTime_Lcl_Done:=FALSE;
bDeter_CondActTime_Clnt_Done:=FALSE;

bStepDone:=FALSE;
IF fbCIP_Source.m_CheckStatus(eReqStatus:=E_CIP_Source.eClose) 
AND fbCIP_Usage.m_CheckStatus(eReqStatus:=E_CIP_Usage.eLocal)  
AND fbCIP_Return.m_CheckStatus(eReqStatus:=E_CIP_Return.eDrain)  
THEN;
	//IF eReq.eClient=E_CIP_Usage.eLocal 
	IF lvlTank_T92.e_state=E_Tank_Level.eLL
	AND lvlTank_T92.rTankLevel>st_CIP_Param.r_Tank92_Volume//st_CIP_Param.r_TankLevel_1//st_CIP_Param.r_Deter_92_TankLvl_1 // Local requered Level
	THEN;	
		bStepDone:=TRUE;
		fbPis.m_SetByRecipe(stPis:=stPis_FillWater_T92, req:=E_Piston_Recipe_State.Release);
	(*ELSIF lvlTank_T92.e_state=E_Tank_Level.eLL
	AND lvlTank_T92.rTankLevel>st_CIP_Param.r_TankVolume_1//Client requered Level
	THEN;
		//Level OK
		bStepDone:=TRUE;
		fbPis.m_SetByRecipe(stPis:=stPis_FillWater_T92, req:=E_Piston_Recipe_State.Release);*)
	ELSE;
		//Fill water
		IF NOT arrTanksSens[E_Tank_Name.T92].get_stTankLevel_OverFlow() THEN;
			fbPis.m_SetByRecipe(stPis:=stPis_FillWater_T92, req:=E_Piston_Recipe_State.Act);			
		END_IF	
	END_IF	
END_IF
END_ACTION

ACTION _aFill_Water_T92_entry:
fbCIP_Source.m_Run(eReqProc:=E_CIP_Source.eClose);
fbCIP_Usage.m_Run(eReqProc:=E_CIP_Usage.eLocal);
fbCIP_Return.m_Run(eReqProc:=E_CIP_Return.eDrain);
bSprinkler:=FALSE;
m_MixProof_set();
m_DashState_activate(stage:=E_CIP_DashStage_List.e03_CIP2_Local_Detergent_Fill);
END_ACTION

ACTION _aFill_Water_T93_active:
bStepDone:=FALSE;
IF fbCIP_Source.m_CheckStatus(eReqStatus:=E_CIP_Source.eClose) 
AND fbCIP_Usage.m_CheckStatus(eReqStatus:=E_CIP_Usage.eLocal)
AND fbCIP_Return.m_CheckStatus(eReqStatus:=E_CIP_Return.eDrain) 
THEN;
	IF TRUE
	AND (lvlTank_T93.e_state=E_Tank_Level.eLL OR TRUE)
	AND lvlTank_T93.rTankLevel>st_CIP_Param.r_Tank93_Volume//fReqVolumeT93 // Client requered Level
	THEN;
		//Level OK
		bStepDone:=TRUE;
		fbPis.m_SetByRecipe(stPis:=stPis_FillWater_T93, req:=E_Piston_Recipe_State.Release);
	ELSE;
		//Fill water
		IF NOT arrTanksSens[E_Tank_Name.T93].get_stTankLevel_OverFlow() THEN;
			fbPis.m_SetByRecipe(stPis:=stPis_FillWater_T93, req:=E_Piston_Recipe_State.Act);			
		END_IF
	END_IF	
	
END_IF
END_ACTION

ACTION _aFill_Water_T93_Done_active:
bStepDone:=FALSE;
IF fbPis.m_CheckByRecipe(stPis:=stPis_FillWater_T93, req:=E_Piston_Recipe_State.Release) THEN
	bStepDone:=TRUE;
END_IF
END_ACTION

ACTION _aFill_Water_T93_Done_entry:
fbPis.m_SetByRecipe(stPis:=stPis_FillWater_T93, req:=E_Piston_Recipe_State.Release);
END_ACTION

ACTION _aFill_Water_T93_entry:
fbCIP_Source.m_Run(eReqProc:=E_CIP_Source.eClose);
fbCIP_Usage.m_Run(eReqProc:=E_CIP_Usage.eLocal);
fbCIP_Return.m_Run(eReqProc:=E_CIP_Return.eDrain);
mCIP_Clients_command(command:=E_CIP_Client_Command.eDrain);



m_DashState_activate(stage:=E_CIP_DashStage_List.e01_CIP1_Client_Drain_Product_Rest_Pipe);
(*
arCIP_DashStage_list[E_CIP_DashStage_List.e01_CIP1_Client_Drain_Product_Rest_Pipe]:=E_CIP_DashStage.eCIPStage_Active;
eCIP_DashStage_actual:=E_CIP_DashStage_List.e01_CIP1_Client_Drain_Product_Rest_Pipe;
sCIP_DashStage_actual:=TO_STRING(eCIP_DashStage_actual);
*)

m_MixProof_set();
END_ACTION

ACTION _aFill_Water_T94_active:
bStepDone:=FALSE;
IF fbCIP_Source.m_CheckStatus(eReqStatus:=E_CIP_Source.eClose) 
AND fbCIP_Usage.m_CheckStatus(eReqStatus:=E_CIP_Usage.eLocal)  
AND fbCIP_Return.m_CheckStatus(eReqStatus:=E_CIP_Return.eDrain)  
THEN;//need something in case there are error in level sensor, should jump into error step and close all valves

	//IF eReq.eClient=E_CIP_Usage.eLocal 
	IF TRUE 
	AND (lvlTank_T94.e_state=E_Tank_Level.eLL OR TRUE)
	AND lvlTank_T94.rTankLevel>st_CIP_Param.r_Tank94_Volume//st_CIP_Param.r_Water_TankLvl_Lcl_1 // Client requered Level
	THEN;	
		bStepDone:=TRUE;
		fbPis.m_SetByRecipe(stPis:=stPis_FillWater_T94, req:=E_Piston_Recipe_State.Release);
	ELSE;
		//Fill water
		IF NOT arrTanksSens[E_Tank_Name.T94].get_stTankLevel_OverFlow() THEN;
			fbPis.m_SetByRecipe(stPis:=stPis_FillWater_T94, req:=E_Piston_Recipe_State.Act);			
		END_IF	END_IF	

END_IF
END_ACTION

ACTION _aFill_Water_T94_Done_active:
bStepDone:=FALSE;
IF fbPis.m_CheckByRecipe(stPis:=stPis_FillWater_T94, 		req:=E_Piston_Recipe_State.Act) THEN
	bStepDone:=TRUE;
END_IF
bStepDone:=TRUE;
END_ACTION

ACTION _aFill_Water_T94_Done_entry:
fbPis.m_SetByRecipe(stPis:=stPis_FillWater_T94, 			req:=E_Piston_Recipe_State.Release);
END_ACTION

ACTION _aFill_Water_T94_entry:
fbCIP_Source.m_Run(eReqProc:=E_CIP_Source.eClose);
fbCIP_Usage.m_Run(eReqProc:=E_CIP_Usage.eLocal);
fbCIP_Return.m_Run(eReqProc:=E_CIP_Return.eDrain);
fbPis.m_SetByRecipe(stPis:=stPis_FillWater_T94, 			req:=E_Piston_Recipe_State.Act);


CASE eRefClient_fbElement.eState_Long OF

	E_Element_State_Long.eCIP_2_Deterged:;
			m_DashState_activate(stage:=E_CIP_DashStage_List.e08_CIP3_Detergent_Collect);

	E_Element_State_Long.eCIP_4_Sanitized:;
			m_DashState_activate(stage:=E_CIP_DashStage_List.e17_CIP5_DisInfection_Collect);
			
END_CASE

m_MixProof_set();
END_ACTION

ACTION _aFlow_Volume_Meter_active:
//

IF eReq.eClient=E_CIP_Usage.eLocal THEN;
	//
ELSE;
	
END_IF

(*

eReq.eClient=E_CIP_Usage.eLocal
*)
END_ACTION

ACTION _aGet_Client_active:
bStepDone:=FALSE;
IF __ISVALIDREF(eRefClient_fbElement) THEN
	IF eRefClient_fbElement.ProdStatus=E_Prod_Status.Active THEN;
		RETURN;
	END_IF
	CASE eReq.eType OF
		E_CIP_Type.R_Water:;
			CASE eRefClient_fbElement.eState_Long OF
				E_Element_State_Long.eNotClean:;
						eRun:=E_CIP_Source.eT93_R_Water;	
			END_CASE
		
		E_CIP_Type.Detergent:;
			CASE eRefClient_fbElement.eState_Long OF
				E_Element_State_Long.eNotClean:;
						eRun:=E_CIP_Source.eT93_R_Water;	
					
				E_Element_State_Long.eCIP_1_Rinzed:;
						eRun:=E_CIP_Source.eT92_Detergent;	
						
				E_Element_State_Long.eCIP_2_Deterged:;
						eRun:=E_CIP_Source.eT94_Water;					
			END_CASE
		
		E_CIP_Type.Full:;
			CASE eRefClient_fbElement.eState_Long OF
				E_Element_State_Long.eNotClean:;
						eRun:=E_CIP_Source.eT93_R_Water;	
					
				E_Element_State_Long.eCIP_1_Rinzed:;
						eRun:=E_CIP_Source.eT92_Detergent;	
					
				E_Element_State_Long.eCIP_2_Deterged:;
						eRun:=E_CIP_Source.eT94_Water;	
					
				E_Element_State_Long.eCIP_3_Deterged_Clean:;
						eRun:=E_CIP_Source.eT91_Sanitation;		
				
				E_Element_State_Long.eCIP_4_Sanitized:;
						eRun:=E_CIP_Source.eT94_Water;					
			END_CASE	
		
	END_CASE
	(*
	IF eRun<>E_CIP_Source.eNone THEN;
		eRefClient_fbElement.m_InterConnect(value:=E_InterConnection.ConnToCIP);
	END_IF	
	*)
	bStepDone:=TRUE;
END_IF
END_ACTION

ACTION _aGet_Client_exit:
m_DashState_ToString_convertion();
m_DashState_Get_ToBeDone_List();
END_ACTION

ACTION _ainit_active:
SFCReset:=FALSE;
END_ACTION

ACTION _ainit_exit:
bRun:=FALSE;
IF eMode=E_CIP_Mode.eAuto THEN;
	eMode:=E_CIP_Mode.eManual;
END_IF
g_Data.b_CIP_Run:=FALSE;
m_MixProof_set();
_aGet_Client_active();
END_ACTION

ACTION _ameasure_Deterg_2_active:

END_ACTION

ACTION _ameasure_Deterg_active:

END_ACTION

ACTION _ameasure_Dis_2_active:

END_ACTION

ACTION _ameasure_Dis_active:

END_ACTION

ACTION _ameasureDelay_CIP2_1_active:
bStepDone:=FALSE;
tMeasureDelayTime:=SECOND_TO_TIME(g_Data.arr_CIP_Param[E_CIP_Usage.eLocal].t_Measure_Delay);
IF measureDelay_CIP2_1.t > tMeasureDelayTime THEN;
	bStepDone:=TRUE;
END_IF

IF bCIP_Condition_Failed THEN;
	bStepDone:=TRUE;
END_IF
END_ACTION

ACTION _ameasureDelay_CIP2_1_entry:
pcDetergent.mReset();
END_ACTION

ACTION _ameasureDelay_CIP2_2_active:
bStepDone:=FALSE;
tMeasureDelayTime:=SECOND_TO_TIME(st_CIP_Param.t_Measure_Delay);
IF measureDelay_CIP2_2.t > tMeasureDelayTime THEN;
	bStepDone:=TRUE;
END_IF

IF bCIP_Condition_Failed THEN;
	bStepDone:=TRUE;
END_IF
END_ACTION

ACTION _ameasureDelay_CIP2_2_entry:
pcDetergent.mReset();
END_ACTION

ACTION _ameasureDelay_CIP3_1_active:
bStepDone:=FALSE;
tMeasureDelayTime:=SECOND_TO_TIME(g_Data.arr_CIP_Param[E_CIP_Usage.eLocal].t_Measure_Delay);
IF measureDelay_CIP3_1.t > tMeasureDelayTime THEN;
	bStepDone:=TRUE;
END_IF

IF bCIP_Condition_Failed THEN;
	bStepDone:=TRUE;
END_IF
END_ACTION

ACTION _ameasureDelay_CIP3_1_entry:
pcDisInfectant.mReset();
END_ACTION

ACTION _ameasureDelay_CIP3_2_active:
bStepDone:=FALSE;
tMeasureDelayTime:= SECOND_TO_TIME(st_CIP_Param.t_Measure_Delay);
IF measureDelay_CIP3_2.t > tMeasureDelayTime 
OR bSprinkler
THEN;
	bStepDone:=TRUE;
END_IF

IF bCIP_Condition_Failed THEN;
	bStepDone:=TRUE;
END_IF
END_ACTION

ACTION _ameasureDelay_CIP3_2_entry:
pcDisInfectant.mReset();
END_ACTION

ACTION _aReady_active:
CASE eMode OF
	E_CIP_Mode.eOff:;
		bRun:=FALSE;
		bStepDone:=FALSE;
	E_CIP_Mode.eManual:;
		IF TRUE 
		AND bRun 
		AND arCIP_RequestBufer[0].eClient<>E_CIP_Usage.eNotInUse
		
		THEN;
			bStepDone:=TRUE;
		ELSE;
			bStepDone:=FALSE;
		END_IF	
	E_CIP_Mode.eAuto:;
		IF TRUE 
		//AND bRun 
		AND arCIP_RequestBufer[0].eClient<>E_CIP_Usage.eNotInUse
		
		THEN;
			bRun:=TRUE;
			bStepDone:=TRUE;
		ELSE;
			bStepDone:=FALSE;
		END_IF		
END_CASE
END_ACTION

ACTION _aReady_exit:
eReq:=arCIP_RequestBufer[0];
bClientTypeIs_Tank:=FALSE;

CASE eReq.eClient OF
	E_CIP_Usage.eLocal:;
		eRefClient_fbElement REF= fbElement_Blank;
		IF eReq.eType=E_CIP_Type.Full THEN;
			eRefClient_fbElement.State:=E_Element_State_Long.eNotClean;
		ELSE;
			eRefClient_fbElement.State:=E_Element_State_Long.eCIP_1_Rinzed;
		END_IF	
		
	E_CIP_Usage.eTank_1:;
		eRefClient_fbElement REF= fbElement[E_Element_List.eTank_1];
		ref_lvlTank_Client REF= stTanksSens[E_Tank_Name.T1];
		bClientTypeIs_Tank:=TRUE;
		
	E_CIP_Usage.eTank_2:;
		eRefClient_fbElement REF= fbElement[E_Element_List.eTank_2];
		ref_lvlTank_Client REF= stTanksSens[E_Tank_Name.T2];
		bClientTypeIs_Tank:=TRUE;
		
	E_CIP_Usage.eTank_3:;
		eRefClient_fbElement REF= fbElement[E_Element_List.eTank_3];
		ref_lvlTank_Client REF= stTanksSens[E_Tank_Name.T3];
		bClientTypeIs_Tank:=TRUE;
		
	E_CIP_Usage.eTank_4:;
		eRefClient_fbElement REF= fbElement[E_Element_List.eTank_4];
		ref_lvlTank_Client REF= stTanksSens[E_Tank_Name.T4];
		bClientTypeIs_Tank:=TRUE;
		
	E_CIP_Usage.eTriBlender_Marinada:;
		eRefClient_fbElement REF= fbElement[E_Element_List.eTriBlender_Marinada];
		
	E_CIP_Usage.eTriBlender_Color:;
		eRefClient_fbElement REF= fbElement[E_Element_List.eTriBlender_Color];
		
	E_CIP_Usage.eLine_Marinada:;
		eRefClient_fbElement REF= fbElement[E_Element_List.eLine_Marinada];
		
	E_CIP_Usage.eLine_Color:;
		eRefClient_fbElement REF= fbElement[E_Element_List.eLine_Color];

END_CASE
g_Data.b_CIP_Run:=TRUE;
bClientRef_done:=TRUE;
m_DashState_MixProof_set();

(*
CASE eCIP_Usage OF
	E_CIP_Usage.eTank_1:;
			IF stTanksSens[E_Tank_Name.T1].e_state=E_Tank_Level.eEmpty THEN;
				bStepDone:=TRUE;	
			END_IF	
	E_CIP_Usage.eTank_2:;
			IF stTanksSens[E_Tank_Name.T2].e_state=E_Tank_Level.eEmpty THEN;
				bStepDone:=TRUE;	
			END_IF	
	E_CIP_Usage.eTank_3:;
			IF stTanksSens[E_Tank_Name.T3].e_state=E_Tank_Level.eEmpty THEN;
				bStepDone:=TRUE;	
			END_IF	
	E_CIP_Usage.eTank_4:;
			IF stTanksSens[E_Tank_Name.T4].e_state=E_Tank_Level.eEmpty THEN;
				bStepDone:=TRUE;	
			END_IF
ELSE;
*)
END_ACTION

ACTION _aReadyToCondition_Count_active:

(*
IF TRUE 
AND pcFlow1_Rate.mRun()
AND pcFlow2_Rate.mRun()
//AND pcPressure.mRun()
THEN;
	bStepDone:=TRUE;
ELSE;
	bStepDone:=FALSE;
END_IF
*)

(*
IF eRefClient_fbElement.eState_Long=E_Element_State_Long.eCIP_2_Deterged THEN;
	
ELSIF eRefClient_fbElement.eState_Long=E_Element_State_Long.eCIP_4_Sanitized THEN;
	
END_IF
*)

(*
IF TRUE //Future condition
AND StartPump_CIP3_02.t>SECOND_TO_TIME(st_CIP_Param.t_PumpInitRun) THEN;
	fb_PumpCIP.m_Run(RPM:=pcFlow1_Rate.mRun_PID(Set_Point:=fFlowRate,controlManual:=NOT(fb_PumpCIP.modeAuto)));
	fb_PumpClient.m_Run(RPM:=st_CIP_Param.r_CIP_Client_Pump);
END_IF
*)
END_ACTION

ACTION _aReadyToCondition_Count_entry:

fb_PumpCIP.m_Run(RPM:=st_CIP_Param.r_CIP_Pump);
fb_PumpClient.m_Run(RPM:=st_CIP_Param.r_CIP_Client_Pump);
END_ACTION

ACTION _aReFill_Water_T93_active:
IF TRUE
//AND lvlTank_T94.e_state=E_Tank_Level.eLL
AND lvlTank_T93.rTankLevel + 0 > st_CIP_Param.r_Tank93_Volume//st_CIP_Param.r_Water_TankLvl_Lcl_1 // Client requered Level
THEN;	
	bStepDone:=TRUE;
	fbPis.m_SetByRecipe(stPis:=stPis_FillWater_T93, req:=E_Piston_Recipe_State.Release);
ELSE;
	//Fill water
	bStepDone:=FALSE;
		IF NOT arrTanksSens[E_Tank_Name.T93].get_stTankLevel_OverFlow() THEN;
			fbPis.m_SetByRecipe(stPis:=stPis_FillWater_T93, req:=E_Piston_Recipe_State.Act);			
		END_IF
END_IF
END_ACTION

ACTION _aReFill_Water_T94_active:
IF TRUE
//AND lvlTank_T94.e_state=E_Tank_Level.eLL
AND lvlTank_T94.rTankLevel +20>st_CIP_Param.r_Tank94_Volume//st_CIP_Param.r_Water_TankLvl_Lcl_1 // Client requered Level
THEN;	
	bStepDone:=TRUE;
	fbPis.m_SetByRecipe(stPis:=stPis_FillWater_T94, req:=E_Piston_Recipe_State.Release);
ELSE;
	//Fill water
	bStepDone:=FALSE;
	IF NOT arrTanksSens[E_Tank_Name.T94].get_stTankLevel_OverFlow() THEN;
		fbPis.m_SetByRecipe(stPis:=stPis_FillWater_T94, req:=E_Piston_Recipe_State.Act);			
	END_IF
END_IF
END_ACTION

ACTION _aReset_Cond_Tm_CIP2_01_active:
tonr_CIP_Condition(ResetTime:=TRUE);
END_ACTION

ACTION _aSet_Valves_ToDeafult_active:
bStepDone:=FALSE;
IF TRUE 
AND fbPis.m_CheckByRecipe(stPis:=stPis_FillWater_T91, 	req:=E_Piston_Recipe_State.Release) 
AND fbPis.m_CheckByRecipe(stPis:=stPis_FillWater_T92, 	req:=E_Piston_Recipe_State.Release) 
AND fbPis.m_CheckByRecipe(stPis:=stPis_FillWater_T93, 	req:=E_Piston_Recipe_State.Release) 
AND fbPis.m_CheckByRecipe(stPis:=stPis_FillWater_T94, 	req:=E_Piston_Recipe_State.Release) 

AND m_MixProof_Release_All()
THEN;
	bStepDone:=TRUE;
END_IF
END_ACTION

ACTION _aSet_Valves_ToDeafult_entry:
fbPis.m_SetByRecipe(stPis:=stPis_FillWater_T91, req:=E_Piston_Recipe_State.Release);
fbPis.m_SetByRecipe(stPis:=stPis_FillWater_T92, req:=E_Piston_Recipe_State.Release);
fbPis.m_SetByRecipe(stPis:=stPis_FillWater_T93, req:=E_Piston_Recipe_State.Release);
fbPis.m_SetByRecipe(stPis:=stPis_FillWater_T94, req:=E_Piston_Recipe_State.Release);

_aDisconnect_n_Drain_CIP_Client_entry();
END_ACTION

ACTION _aSprinkler_Request_CIP1_active:


IF TRUE // Type Tank
AND bClientTypeIs_Tank	
AND bSprinkler
THEN;	
	bStepDone:=TRUE;
	m_DashState_done(stage:=E_CIP_DashStage_List.e02_CIP1_Client_Drain_Product_Rest_Sprinkler);
	
ELSIF TRUE // Type Pine
AND NOT bClientTypeIs_Tank	
THEN;	
	bStepDone:=TRUE;
	m_DashState_done(stage:=E_CIP_DashStage_List.e01_CIP1_Client_Drain_Product_Rest_Pipe);
	
ELSE;
	//continue with sprinkler
	bStepDone:=FALSE;
	m_DashState_done(stage:=E_CIP_DashStage_List.e01_CIP1_Client_Drain_Product_Rest_Pipe);
	m_DashState_activate(stage:=E_CIP_DashStage_List.e02_CIP1_Client_Drain_Product_Rest_Sprinkler);
	
END_IF
END_ACTION

ACTION _aSprinkler_Request_CIP4_active:


IF TRUE // Type Tank
AND bClientTypeIs_Tank	
AND bSprinkler
THEN;	
	bStepDone:=TRUE;
	CASE eRefClient_fbElement.eState_Long OF
	
		E_Element_State_Long.eCIP_2_Deterged:;
				m_DashState_done(stage:=E_CIP_DashStage_List.e11_CIP3_Detergent_Clean_Sprinkler);
	
		E_Element_State_Long.eCIP_4_Sanitized:;
				m_DashState_done(stage:=E_CIP_DashStage_List.e20_CIP5_DisInfection_Clean_Sprinkler);
				
	END_CASE	
	
ELSIF TRUE // Type Pine
AND NOT bClientTypeIs_Tank	
THEN;	
	bStepDone:=TRUE;
	CASE eRefClient_fbElement.eState_Long OF
	
		E_Element_State_Long.eCIP_2_Deterged:;
				m_DashState_done(stage:=E_CIP_DashStage_List.e10_CIP3_Detergent_Clean_Pipe);
	
		E_Element_State_Long.eCIP_4_Sanitized:;
				m_DashState_done(stage:=E_CIP_DashStage_List.e19_CIP5_DisInfection_Clean_Pipe);
				
	END_CASE	
	
ELSE;
	//continue with sprinkler
	bStepDone:=FALSE;
	CASE eRefClient_fbElement.eState_Long OF
	
		E_Element_State_Long.eCIP_2_Deterged:;
				m_DashState_done(stage:=E_CIP_DashStage_List.e10_CIP3_Detergent_Clean_Pipe);
				m_DashState_activate(stage:=E_CIP_DashStage_List.e11_CIP3_Detergent_Clean_Sprinkler);
	
		E_Element_State_Long.eCIP_4_Sanitized:;
				m_DashState_done(stage:=E_CIP_DashStage_List.e19_CIP5_DisInfection_Clean_Pipe);
				m_DashState_activate(stage:=E_CIP_DashStage_List.e20_CIP5_DisInfection_Clean_Sprinkler);
				
	END_CASE	
	
END_IF
END_ACTION

ACTION _aStartPump_CIP1_01_active:
bStepDone:=FALSE;
(*
IF StartPump_CIP1_01.t>SECOND_TO_TIME(st_CIP_Param.t_PumpInitRun) 
OR lvlTank_T93.rTankLevel<st_CIP_Param.r_Tank93_Volume//st_CIP_Param.r_RWater_93_TankLvl
THEN//Time+flow+water volume
	bStepDone:=TRUE;
END_IF
*)
bStepDone:=TRUE;
END_ACTION

ACTION _aStartPump_CIP1_01_entry:
fb_PumpCIP.m_Run(RPM:=st_CIP_Param.r_CIP_Pump);
fb_PumpClient.m_Run(RPM:=st_CIP_Param.r_CIP_Client_Pump);

mVolumeReset_All();

tonr_CIP_Condition(ResetTime:=TRUE);
END_ACTION

ACTION _aStartPump_CIP2_01_active:
IF TRUE 
//AND stAnalogSensor[E_ASense_Name.FT1001].Value>=g_Data.arr_CIP_Param[E_CIP_Usage.eLocal].r_Flow_1 // 
//AND stAnalogSensor[E_ASense_Name.FT1002].Value>=g_Data.arr_CIP_Param[E_CIP_Usage.eLocal].r_Flow_2 // 
//AND stAnalogSensor[E_ASense_Name.PT1001].Value>=g_Data.arr_CIP_Param[E_CIP_Usage.eLocal].r_Pressure // 
//AND pcFlow1_Rate.mRun_With_SP(Set_Point:=g_Data.arr_CIP_Param[E_CIP_Usage.eLocal].r_Flow_Pipe)
//AND pcFlow2_Rate.mRun_With_SP(Set_Point:=g_Data.arr_CIP_Param[E_CIP_Usage.eLocal].r_Flow_Pipe)
AND pcFlow1_Rate.mRun()
AND pcFlow2_Rate.mRun()
//AND pcPressure.mRun()
THEN;
	bStepDone:=TRUE;
ELSE;
	bStepDone:=FALSE;
END_IF

fb_PumpCIP.m_Run(RPM:=pcFlow1_Rate.mRun_PID(Set_Point:=g_Data.arr_CIP_Param[E_CIP_Usage.eLocal].r_Flow_Pipe,controlManual:=NOT(fb_PumpCIP.modeAuto)));
END_ACTION

ACTION _aStartPump_CIP2_01_entry:

//fb_PumpDetergent.m_Auto();
fb_HeatExchenger.m_Auto();
bCIP_Condition_Failed:=FALSE;
bCIP_Condition_Done:=FALSE;
iConcentrationDeluteCounter:=0;

nStepHeat:=1;
END_ACTION

ACTION _aStartPump_CIP2_02_active:
fb_PumpCIP.m_Run(RPM:=pcFlow1_Rate.mRun_PID(Set_Point:=fFlowRate, controlManual:=NOT(fb_PumpCIP.modeAuto)));
fb_PumpClient.m_Run(RPM:=st_CIP_Param.r_CIP_Client_Pump);

IF TRUE 
AND pcFlow1_Rate.mRun()
AND pcFlow2_Rate.mRun()
//AND pcPressure.mRun()
THEN;
	bStepDone:=TRUE;
ELSE;
	bStepDone:=FALSE;
END_IF
END_ACTION

ACTION _aStartPump_CIP2_02_entry:
fb_HeatExchenger.m_Auto();
bCIP_Condition_Failed:=FALSE;
bCIP_Condition_Done:=FALSE;
iConcentrationDeluteCounter:=0;

nStepHeat:=10;
END_ACTION

ACTION _aStartPump_CIP2_RPM_01_active:
bStepDone:=FALSE;
fb_PumpCIP.m_Run(RPM:=g_Data.arr_CIP_Param[E_CIP_Usage.eLocal].r_CIP_Pump);//1500

IF TRUE //Future condition
AND StartPump_CIP2_RPM_01.t>SECOND_TO_TIME(g_Data.arr_CIP_Param[E_CIP_Usage.eLocal].t_PumpInitRun) 
AND fb_PumpCIP.nRPM=g_Data.arr_CIP_Param[E_CIP_Usage.eLocal].r_CIP_Pump
//AND stAnalogSensor[E_ASense_Name.FT1001].Value>=g_Data.arr_CIP_Param[E_CIP_Usage.eLocal].r_Flow_Pipe // 
//AND stAnalogSensor[E_ASense_Name.FT1002].Value>=g_Data.arr_CIP_Param[E_CIP_Usage.eLocal].r_Flow_Pipe // 
THEN;
	bStepDone:=TRUE;
END_IF
END_ACTION

ACTION _aStartPump_CIP2_RPM_02_active:
bStepDone:=FALSE;

fb_PumpCIP.m_Run(RPM:=st_CIP_Param.r_CIP_Pump);
fb_PumpClient.m_Run(RPM:=st_CIP_Param.r_CIP_Client_Pump);
bStepDone:=TRUE;

// to stas question ? deference:
//fb_PumpCIP.m_Run(RPM:=g_Data.arr_CIP_Param[E_CIP_Usage.eLocal].r_CIP_Pmp_1);//1500
//fb_PumpCIP.m_Run(RPM:=st_CIP_Param.r_CIP_Pmp_1);
(*
IF TRUE //Future condition
AND delta_T92_Volume < - st_CIP_Param.r_Volume_Solution_Fill // Volume 
//AND StartPump_CIP2_RPM_02.t>SECOND_TO_TIME(g_Data.arr_CIP_Param[E_CIP_Usage.eLocal].t_PumpInitRun) 
THEN;
	bStepDone:=TRUE;
END_IF
*)
END_ACTION

ACTION _aStartPump_CIP2_RPM_02_entry:
mVolumeReset_All();
tonr_CIP_Condition(ResetTime:=TRUE);
END_ACTION

ACTION _aStartPump_CIP2_RPM_03_active:
bStepDone:=FALSE;
fb_PumpCIP.m_Run(RPM:=g_Data.arr_CIP_Param[E_CIP_Usage.eLocal].r_CIP_Pump);

IF TRUE //Future condition
AND StartPump_CIP2_RPM_03.t>SECOND_TO_TIME(g_Data.arr_CIP_Param[E_CIP_Usage.eLocal].t_PumpInitRun) 
THEN;
	bStepDone:=TRUE;
END_IF
END_ACTION

ACTION _aStartPump_CIP2_RPM_04_active:
bStepDone:=FALSE;
fb_PumpCIP.m_Run(RPM:=pcFlow1_Rate.mRun_PID(Set_Point:=st_CIP_Param.r_CIP_Pump,controlManual:=NOT(fb_PumpCIP.modeAuto)));
fb_PumpClient.m_Run(RPM:=st_CIP_Param.r_CIP_Client_Pump);

IF TRUE //Future condition
AND StartPump_CIP2_RPM_04.t>SECOND_TO_TIME(st_CIP_Param.t_PumpInitRun) 
THEN;
	bStepDone:=TRUE;
END_IF
END_ACTION

ACTION _aStartPump_CIP3_01_active:
IF TRUE 
(*AND stAnalogSensor[E_ASense_Name.FT1001].Value>=g_Data.arr_CIP_Param[E_CIP_Usage.eLocal].r_Flow_1//200 // 
AND stAnalogSensor[E_ASense_Name.FT1002].Value>=g_Data.arr_CIP_Param[E_CIP_Usage.eLocal].r_Flow_2//200 // 
AND stAnalogSensor[E_ASense_Name.PT1001].Value>=g_Data.arr_CIP_Param[E_CIP_Usage.eLocal].r_Pressure//0.5 //*)
AND pcFlow1_Rate.mRun()
AND pcFlow2_Rate.mRun()
//AND pcPressure.mRun()
THEN;
	bStepDone:=TRUE;
ELSE;
	bStepDone:=FALSE;
END_IF

fb_PumpCIP.m_Run(RPM:=pcFlow1_Rate.mRun_PID(Set_Point:=g_Data.arr_CIP_Param[E_CIP_Usage.eLocal].r_Flow_Pipe,controlManual:=NOT(fb_PumpCIP.modeAuto)));
END_ACTION

ACTION _aStartPump_CIP3_01_entry:


fb_HeatExchenger.m_Auto();
bCIP_Condition_Failed:=FALSE;
bCIP_Condition_Done:=FALSE;

nStepHeat:=2;
iConcentrationDeluteCounter:=0;
END_ACTION

ACTION _aStartPump_CIP3_02_active:
IF TRUE 
(*AND stAnalogSensor[E_ASense_Name.FT1001].Value>=st_CIP_Param.r_Flow_1 // 
AND stAnalogSensor[E_ASense_Name.FT1002].Value>=st_CIP_Param.r_Flow_2 // 
AND stAnalogSensor[E_ASense_Name.PT1001].Value>=st_CIP_Param.r_Pressure // *)
AND pcFlow1_Rate.mRun()
AND pcFlow2_Rate.mRun()
//AND pcPressure.mRun()
THEN;
	bStepDone:=TRUE;
ELSE;
	bStepDone:=FALSE;
END_IF

//fb_PumpCIP.m_Run(RPM:=pcFlow1_Rate.mRun_PID(Set_Point:=fFlowRate,controlManual:=NOT(fb_PumpCIP.modeAuto)));
//fb_PumpClient.m_Run(RPM:=pcFlow2_Rate.mRun_PID(Set_Point:=fFlowRate,controlManual:=NOT(fb_PumpCIP.modeAuto)));

IF TRUE //Future condition
AND StartPump_CIP3_02.t>SECOND_TO_TIME(st_CIP_Param.t_PumpInitRun) THEN;
	fb_PumpCIP.m_Run(RPM:=pcFlow1_Rate.mRun_PID(Set_Point:=fFlowRate,controlManual:=NOT(fb_PumpCIP.modeAuto)));
	fb_PumpClient.m_Run(RPM:=st_CIP_Param.r_CIP_Client_Pump);
END_IF

IF NOT bSprinkler THEN
	//pipe
	tConditionTime	:=st_CIP_Param.t_ConditionDisInfection;
	fFlowRate		:=st_CIP_Param.r_Flow_Pipe;
	//rVolume_Collect :=st_CIP_Param.r_Volume_Collect_DisInfection;
	//rVolume_Drain	:=st_CIP_Param.r_Volume_Drain_DisInfection;
	//rVolume_Recycle	:=st_CIP_Param.r_Volume_Recycle_DisInfection;
ELSE
	//sprinkler
	tConditionTime	:=st_CIP_Param.t_ConditionDisInfection_Sprinkler;
	fFlowRate		:=st_CIP_Param.r_Flow_Sprinkler;
	//rVolume_Collect :=st_CIP_Param.r_Volume_Collect_DisInfection*st_CIP_Param.r_Volume_Sprinkler_Ratio;
	//rVolume_Drain	:=st_CIP_Param.r_Volume_Drain_DisInfection*st_CIP_Param.r_Volume_Sprinkler_Ratio;
	//rVolume_Recycle	:=st_CIP_Param.r_Volume_Recycle_DisInfection*st_CIP_Param.r_Volume_Sprinkler_Ratio;
END_IF
END_ACTION

ACTION _aStartPump_CIP3_02_entry:
(*fb_PumpCIP.m_Run(RPM:=st_CIP_Param.r_CIP_Pmp_1);
fb_PumpClient.m_Run(RPM:=st_CIP_Param.r_CIP_Client_Pmp_1);*)
//fb_PumpDisinfection.m_Auto();
	
//Heat Exchenger	
fb_HeatExchenger.m_Auto();

bCIP_Condition_Failed:=FALSE;
bCIP_Condition_Done:=FALSE;
iConcentrationDeluteCounter:=0;

nStepHeat:=20;
END_ACTION

ACTION _aStartPump_CIP4_active:
bStepDone:=FALSE;
IF TRUE 
//AND fbPis.m_CheckByRecipe(stPis:=stPis_FillWater_T94, 		req:=E_Piston_Recipe_State.NoChanges) 
THEN
	//bStepDone:=TRUE;
END_IF
bStepDone:=TRUE;
END_ACTION

ACTION _aStartPump_CIP4_entry:
//fbPis.m_SetByRecipe(stPis:=stPis_FillWater_T94, 	req:=E_Piston_Recipe_State.NoChanges);
fb_PumpCIP.m_Run(RPM:=st_CIP_Param.r_CIP_Pump);
fb_PumpClient.m_Run(RPM:=st_CIP_Param.r_CIP_Client_Pump);

mVolumeReset_All();
bSprinkler:=FALSE;
tonr_CIP_Condition(ResetTime:=TRUE);
END_ACTION

ACTION _aStop_Pump_entry:
fb_PumpCIP.m_Stop();
fb_PumpClient.m_Stop();
fb_Stirrer.m_Stop();
fb_PumpDetergent.m_Stop();
fb_PumpDisinfection.m_Stop();
END_ACTION

ACTION _aStopPump_CIP1_01_entry:
fb_PumpCIP.m_Stop();
END_ACTION

ACTION _aStopPump_CIP1_02_entry:
fb_PumpCIP.m_Stop();
fb_PumpClient.m_Stop();
END_ACTION

ACTION _aStopPump_CIP2_01_entry:
fb_PumpCIP.m_Stop();

m_DashState_done(stage:=E_CIP_DashStage_List.e04_CIP2_Local_Detergent_Condition);
END_ACTION

ACTION _aStopPump_CIP2_02_entry:
fb_PumpCIP.m_Stop();
END_ACTION

ACTION _aStopPump_CIP2_03_entry:
fb_PumpCIP.m_Stop();
END_ACTION

ACTION _aStopPump_CIP3_01_entry:
fb_PumpCIP.m_Stop();

m_DashState_done(stage:=E_CIP_DashStage_List.e13_CIP4_Local_DisInfection_Condition);
END_ACTION

ACTION _aStopPump_CIP3_02_entry:
fb_PumpCIP.m_Stop();
END_ACTION

ACTION _aStopPump_CIP3_03_entry:
fb_PumpCIP.m_Stop();
END_ACTION

ACTION _aStopPump_CIP4_01_entry:
fb_PumpCIP.m_Stop();
END_ACTION

ACTION _aStopPump_CIP4_02_entry:
fb_PumpCIP.m_Stop();
fb_PumpClient.m_Stop();
END_ACTION

ACTION _aTank_LowLevel_CIP1_01_active:
bStepDone:=m_Check_ProductionTank_Low_Level();
END_ACTION

ACTION _aTank_LowLevel_CIP1_02_active:
bStepDone:=m_Check_ProductionTank_Low_Level();
END_ACTION

ACTION _aTank_LowLevel_CIP1_02_entry:
fb_PumpCIP.m_Stop();
END_ACTION

ACTION _aTank_LowLevel_CIP2_01_active:
bStepDone:=m_Check_ProductionTank_Low_Level();
END_ACTION

ACTION _aTank_LowLevel_CIP2_02_active:
bStepDone:=m_Check_ProductionTank_Low_Level();
END_ACTION

ACTION _aTank_LowLevel_CIP2_02_entry:
fb_PumpCIP.m_Stop();
fb_PumpClient.m_Run(RPM:=st_CIP_Param.r_CIP_Client_Pump);
END_ACTION

ACTION _aTank_LowLevel_CIP3_01_active:
bStepDone:=m_Check_ProductionTank_Low_Level();
END_ACTION

ACTION _aTank_LowLevel_CIP3_02_active:
bStepDone:=m_Check_ProductionTank_Low_Level();
END_ACTION

ACTION _aTank_LowLevel_CIP3_02_entry:
fb_PumpCIP.m_Stop();
fb_PumpClient.m_Run(RPM:=st_CIP_Param.r_CIP_Client_Pump);
END_ACTION

ACTION _aTank_LowLevel_CIP4_01_active:
bStepDone:=m_Check_ProductionTank_Low_Level();
END_ACTION

ACTION _aTank_LowLevel_CIP4_02_active:
bStepDone:=m_Check_ProductionTank_Low_Level();
END_ACTION

ACTION _aTank_LowLevel_CIP4_02_entry:
fb_PumpCIP.m_Stop();
END_ACTION

ACTION _aTank_MixProof_Clean_CIP2_active:
m_MixProof_run();

IF bValveCleanDone THEN;
	bStepDone:=TRUE;	
ELSE;
	bStepDone:=FALSE;
END_IF
END_ACTION

ACTION _aTank_MixProof_Clean_CIP2_entry:
fb_PumpCIP.m_Stop();
END_ACTION

ACTION _aTank_MixProof_Clean_CIP3_active:
m_MixProof_run();

IF bValveCleanDone THEN;
	bStepDone:=TRUE;	
ELSE;
	bStepDone:=FALSE;
END_IF
END_ACTION

ACTION _aTank_MixProof_Clean_CIP3_entry:
fb_PumpCIP.m_Stop();
END_ACTION

ACTION _aTriBlender_Selection_active:

IF eRefClient_fbElement.eElementID=E_Element_List.eTriBlender_Marinada THEN;
	bStepDone:=fbTriBlender_Select.m_CheckStatus(eReqStatus:=E_TriBlenderSelect.eMarinade);

ELSIF eRefClient_fbElement.eElementID=E_Element_List.eTriBlender_Color THEN;
	bStepDone:=fbTriBlender_Select.m_CheckStatus(eReqStatus:=E_TriBlenderSelect.eColor);
	
ELSE;
	bStepDone:=TRUE;
END_IF
END_ACTION

ACTION _aTriBlender_Selection_entry:

IF eRefClient_fbElement.eElementID=E_Element_List.eTriBlender_Marinada THEN;
	fbTriBlender_Select.m_Run(eReqProc:=E_TriBlenderSelect.eMarinade);
END_IF

IF eRefClient_fbElement.eElementID=E_Element_List.eTriBlender_Color THEN;
	fbTriBlender_Select.m_Run(eReqProc:=E_TriBlenderSelect.eColor);
END_IF
END_ACTION

ACTION _aWaiting_Client_Drain_Done_active:
_aDisconnect_n_Drain_CIP_Client_active();
END_ACTION

ACTION act_CallProcessControl:
//Heat Exchanger
	stHeatExchanger.rValue:=g_AnalogSensor.stAnalogSensor[E_ASense_Name.TT1105].Value;
	//stHeatExchanger.rSetPoint:=st_CIP_Param.r_Temper_ClientReturn;
	pcHeatExchanger(stProcessControl:=stHeatExchanger );
//Client temperature return
	stTemp_ClntReturn.rValue:=g_AnalogSensor.stAnalogSensor[E_ASense_Name.TT1101].Value;//gIO.fbScaleFactor[E_ASense_Name.TT1101].rValOut;
	//stTemp_ClntReturn.rSetPoint:=st_CIP_Param.n _ClientReturn;
	pcTemp_ClntReturn(stProcessControl:=stTemp_ClntReturn );

//Detergent
	//Concentration
	stDetergent.rValue:=g_AnalogSensor.stAnalogSensor[E_ASense_Name.CT1101_3].Value;
	//###stDetergent.ToleranceHigh:=0.05;
	//###stDetergent.ToleravceLow:=0.05;
	//###stDetergent.rSetPoint:=st_CIP_Param.r_DetergentConcentration;//0.3;
	pcDetergent(stProcessControl:=stDetergent );
		
	//Temperature
	//stTemperature_Deterg.rValue:=testTemperature;
	stTemperature_Deterg.rValue:=g_AnalogSensor.stAnalogSensor[E_ASense_Name.TT1003].Value;
	//###stTemperature_Deterg.ToleranceHigh:=1;
	//###stTemperature_Deterg.ToleravceLow:=1;
	//###stTemperature_Deterg.rSetPoint:=st_CIP_Param.r_Temper_Detergent;
	pcTemperature_Deterg(stProcessControl:=stTemperature_Deterg );


//Disinfectant
	//Concentration
	stDisInfectant.rValue:=g_AnalogSensor.stAnalogSensor[E_ASense_Name.CT1101_4].Value;
	//###stDisInfectant.ToleranceHigh:=0.05;
	//###stDisInfectant.ToleravceLow:=0.05;
	//###stDisInfectant.rSetPoint:=st_CIP_Param.r_DisInfectionConcentration;//0.3;
	pcDisInfectant(stProcessControl:=stDisInfectant );
		
	//Temperature	
	//stTemperature_Dis.rValue:=testTemperature;
	stTemperature_Dis.rValue:=g_AnalogSensor.stAnalogSensor[E_ASense_Name.TT1004].Value;
	//###stTemperature_Dis.ToleranceHigh:=1;//0.5
	//###stTemperature_Dis.ToleravceLow:=1;//0.5
	//###stTemperature_Dis.rSetPoint:=st_CIP_Param.r_Temper_DisInfection;//65;
	pcTemperature_Dis(stProcessControl:=stTemperature_Dis );	
	
// Flow_Rate
	//CIP Pump
		//Pump CIP infeed
		stFlow1_Rate.rValue:=g_AnalogSensor.stAnalogSensor[E_ASense_Name.FT1001].Value;
		stFlow1_Rate.rValue:=g_AnalogSensor.stAnalogSensor[E_ASense_Name.FT1001].Value;
		stFlow1_Rate.rValue_Min_To_ReleaseControl:=50;// Litter/Hours
		//stFlow1_Rate.rSetPoint:=st_CIP_Param.r_Flow_Pipe;//:=150
		stFlow1_Rate.bPause:=stOper[E_ModeZone.eCIP].iActOperation=E_OperationButtons.ePauseAll;
		stFlow1_Rate.fCtrlOutput_Manual:=fb_PumpCIP.nRPM;
		stFlow1_Rate.fCtrlOutput_Max:=1700;
		stFlow1_Rate.fCtrlOutput_Min:=700;
		pcFlow1_Rate(stProcessControl:=stFlow1_Rate, );

		//Pump CIP return 
		stFlow2_Rate.rValue:=g_AnalogSensor.stAnalogSensor[E_ASense_Name.FT1002].Value;
		stFlow3_Rate.rValue:=g_AnalogSensor.stAnalogSensor[E_ASense_Name.FT1002].Value;
		stFlow3_Rate.rSetPoint:=stFlow2_Rate.rSetPoint;
		pcFlow2_Rate(stProcessControl:=stFlow2_Rate );
		pcFlow3_Rate(stProcessControl:=stFlow3_Rate );

		// TBD : to check if the first loop(local prepare) when Client selected gets relevant Flow SetPoint 
		IF bSprinkler THEN
			stFlow1_Rate.rSetPoint:=st_CIP_Param.r_Flow_Sprinkler;
			stFlow2_Rate.rSetPoint:=st_CIP_Param.r_Flow_Sprinkler;
		ELSE
			stFlow1_Rate.rSetPoint:=st_CIP_Param.r_Flow_Pipe;
			stFlow2_Rate.rSetPoint:=st_CIP_Param.r_Flow_Pipe;
		END_IF		
		
	//CIP Client Color pump
		//stColor_Level.rValue:=g_AnalogSensor.stAnalogSensor[E_ASense_Name.LT4002].Value;
		stColor_Level.rValue:=g_AnalogSensor.stAnalogSensor[E_ASense_Name.LT4001].Value;
		//###stColor_Level.ToleranceHigh:=10;
		//###stColor_Level.ToleravceLow:=10;
		//stFlow_Rate.rSetPoint:=150;
		pcColor_Level(stProcessControl:=stColor_Level );
	//CIP Client Marinada pump
		stMarinada_Level.rValue:=g_AnalogSensor.stAnalogSensor[E_ASense_Name.LT3002].Value;
		//###stMarinada_Level.ToleranceHigh:=10;
		//###stMarinada_Level.ToleravceLow:=10;
		//stFlow_Rate.rSetPoint:=150;
		pcMarinada_Level(stProcessControl:=stMarinada_Level );
		
//Presure
		stP1001_Pressure.rValue:=g_AnalogSensor.stAnalogSensor[E_ASense_Name.PT1001].Value;
		pcP1001_Pressure(stProcessControl:=stP1001_Pressure );
(*		
		stP3001_Pressure.rValue:=g_AnalogSensor.stAnalogSensor[E_ASense_Name.PT3001].Value;
		pcP3001_Pressure(stProcessControl:=stP3001_Pressure );
		
		stP3002_Pressure.rValue:=g_AnalogSensor.stAnalogSensor[E_ASense_Name.PT3002].Value;
		pcP3002_Pressure(stProcessControl:=stP3002_Pressure );
		
		stP4001_Pressure.rValue:=g_AnalogSensor.stAnalogSensor[E_ASense_Name.PT4001].Value;
		pcP4001_Pressure(stProcessControl:=stP4001_Pressure );
		
		stP4002_Pressure.rValue:=g_AnalogSensor.stAnalogSensor[E_ASense_Name.PT4002].Value;
		pcP4002_Pressure(stProcessControl:=stP4002_Pressure );
			
//TriBlender Flow
		stTriBlender_Flow.rValue:=g_AnalogSensor.stAnalogSensor[E_ASense_Name.FT9011].Value;
		pcTriBlender_Flow(stProcessControl:=stTriBlender_Flow );

//Color skid Concentration
		stColor_TriB_Conc.rValue:=g_AnalogSensor.stAnalogSensor[E_ASense_Name.CT4101].Value;
		pcColor_TriB_Conc(stProcessControl:=stColor_TriB_Conc );		

		stColor_Line_Conc.rValue:=g_AnalogSensor.stAnalogSensor[E_ASense_Name.CT4101].Value;
		pcColor_Line_Conc(stProcessControl:=stColor_Line_Conc );		
*)

//Load def set points
IF bLoadDefSetPoints THEN
	bLoadDefSetPoints:=FALSE;
	mLoadDefProcessSetPoints();
END_IF
		
//selecting set point based on user
	
	IF bTestPID THEN;
		pcFlow1_Rate.mRun();
		pcColor_Level.mRun();

		fb_PumpCIP.m_Auto(control:=pcFlow1_Rate.mRun_PID(Set_Point:=180,controlManual:=NOT(fb_PumpCIP.modeAuto)));
		
		//by CIP Pump RPM control		
		g_Pump.fbPump[E_Pump_List.P4002].m_Auto(control:=pcColor_Level.mRun_Hyst());
		
		IF fb_PumpCIP.modeAuto THEN;
			stFlow1_Rate.bManual:=FALSE;
		ELSE;
			stFlow1_Rate.bManual:=TRUE;
			stFlow1_Rate.fCtrlOutput_Manual:=fb_PumpCIP.nRPM;
		END_IF
		
		IF fb_PumpClient.modeAuto THEN;
			stColor_Level.bManual:=FALSE;
		ELSE;
			stColor_Level.bManual:=TRUE;
			stColor_Level.fCtrlOutput_Manual:=g_Pump.fbPump[E_Pump_List.P4002].nRPM;//fb_PumpClient.nRPM;
		END_IF
			
	END_IF
END_ACTION

ACTION act_GetReference:
stPis_FillWater_T91 REF= stPis[valFillWater_T91];
stPis_FillWater_T92 REF= stPis[valFillWater_T92];
stPis_FillWater_T93 REF= stPis[valFillWater_T93];
stPis_FillWater_T94 REF= stPis[valFillWater_T94];

	//concentration
stDetergent 	REF=g_ProcControl.arr_stProcCntrl[E_ProcessControl_Name.eDetergentConc];
pcDetergent 	REF=g_ProcControl.arr_fbProcCntrl[E_ProcessControl_Name.eDetergentConc];

stDisInfectant 	REF=g_ProcControl.arr_stProcCntrl[E_ProcessControl_Name.eDisinfectionConc];
pcDisInfectant 	REF=g_ProcControl.arr_fbProcCntrl[E_ProcessControl_Name.eDisinfectionConc];

	//Temperature
stTemperature_Deterg REF=g_ProcControl.arr_stProcCntrl[E_ProcessControl_Name.eDeterTemp];
pcTemperature_Deterg REF=g_ProcControl.arr_fbProcCntrl[E_ProcessControl_Name.eDeterTemp];

stTemperature_Dis 	 REF=g_ProcControl.arr_stProcCntrl[E_ProcessControl_Name.eDisTemp];
pcTemperature_Dis 	 REF=g_ProcControl.arr_fbProcCntrl[E_ProcessControl_Name.eDisTemp];
	//Flow rate
stFlow1_Rate REF=g_ProcControl.arr_stProcCntrl[E_ProcessControl_Name.eCIP_Flow_1];
pcFlow1_Rate REF=g_ProcControl.arr_fbProcCntrl[E_ProcessControl_Name.eCIP_Flow_1];

stFlow2_Rate REF=g_ProcControl.arr_stProcCntrl[E_ProcessControl_Name.eCIP_Flow_2];
pcFlow2_Rate REF=g_ProcControl.arr_fbProcCntrl[E_ProcessControl_Name.eCIP_Flow_2];

stFlow3_Rate REF=g_ProcControl.arr_stProcCntrl[E_ProcessControl_Name.eCIP_Flow_3];
pcFlow3_Rate REF=g_ProcControl.arr_fbProcCntrl[E_ProcessControl_Name.eCIP_Flow_3];

	//Level
stColor_Level    REF=g_ProcControl.arr_stProcCntrl[E_ProcessControl_Name.eColor_Level];
pcColor_Level    REF=g_ProcControl.arr_fbProcCntrl[E_ProcessControl_Name.eColor_Level];

stMarinada_Level REF=g_ProcControl.arr_stProcCntrl[E_ProcessControl_Name.eMarin_Level];
pcMarinada_Level REF=g_ProcControl.arr_fbProcCntrl[E_ProcessControl_Name.eMarin_Level];
	//Pressure
stP1001_Pressure 	REF=g_ProcControl.arr_stProcCntrl[E_ProcessControl_Name.eCIP_Pressure];
pcP1001_Pressure 	REF=g_ProcControl.arr_fbProcCntrl[E_ProcessControl_Name.eCIP_Pressure];

//temperature control
stTemp_ClntReturn REF=g_ProcControl.arr_stProcCntrl[E_ProcessControl_Name.eClientReturn_Temp];
pcTemp_ClntReturn REF=g_ProcControl.arr_fbProcCntrl[E_ProcessControl_Name.eClientReturn_Temp];

stHeatExchanger REF=g_ProcControl.arr_stProcCntrl[E_ProcessControl_Name.eHeatExchanger];
pcHeatExchanger REF=g_ProcControl.arr_fbProcCntrl[E_ProcessControl_Name.eHeatExchanger];
END_ACTION

ACTION act_HeatExchng:
//calling heat exchanger 
fb_HeatExchenger(stHeatExchanger:=g_Data.stHeatExchanger );

//Choosing heat exchanger set point 

